(* Logix 5000 project; controller TFF vendor 1 type 14 code 107 rev 34.11; software revision 34.03; part 7 of 36 *)

        [24]   // Product Recovery 1&5 - Empty Recycle Bag (TF3S)
        [16]   // Recycle Bag Fill
        [6]   // Buffer Source Open
        [25]   // Product Recovery 2 - Empty Membranes (TF3S
        [30]   // Filter User
        [34]   // Column User
        [36]   // Fraction 3
        [37]   // Fraction 2
        [61]   // Reserved : Open All valves
        [38]   // Fraction 1
        [18]   // Recovery Filter Flush
        [39]   // System Drain
        [19]   // Batch UF or Membrane Recycle
        [14]   // Membrane Soak
        [2]   // Critical Alarm Flowpath
        [33]   // Column Bypass
        [9]   // Air Source Open
        [4]   // All Source Valves Closed
        [62]   // Reserved : Close All valves
        [3]   // All Source Valves Open
        [8]   // Water Source Open
        [22]   // Product Recovery 2 - Empty Retentate Line (TF2S)
        [26]   // Product Recovery 3&6 - Empty Bypass (TF3S)
        [27]   // Product Recovery 4 - Empty Retentate Line (TF3S)
   FlowPath_Storage : FlowPath[6,64] := ([0,0].Truth1 := -1, [0,0].Mask1 := -1, [0,0].Desc := 'Reserved', [0,1].Status := 1, [0,1].Truth1 := 2097151, [0,1].Mask1 := -1, [0,1].Desc := 'Default', [0,2].Status := 1, [0,2].Truth1 := 539146240, [0,2].Mask1 := -1, [0,2].Desc := 'Critical', [0,3].Status := 1, [0,3].Mask1 := 2047, [0,3].Desc := 'Close All Inlets', [0,4].Truth1 := 17, [0,4].Mask1 := 63, [0,4].Desc := 'Inlet 1A', [0,5].Truth1 := 18, [0,5].Mask1 := 63, [0,5].Desc := 'Inlet 1B', [0,6].Truth1 := 20, [0,6].Mask1 := 63, [0,6].Desc := 'Inlet 1C', [0,7].Truth1 := 24, [0,7].Mask1 := 63, [0,7].Desc := 'Inlet 1D', [0,8].Truth1 := 32, [0,8].Mask1 := 63, [0,8].Desc := 'Inlet 1E', [0,9].Truth1 := 64, [0,9].Mask1 := 1984, [0,9].Desc := 'Inlet 2A', [0,10].Truth1 := 128, [0,10].Mask1 := 1984, [0,10].Desc := 'Inlet 2B', [0,11].Truth1 := 256, [0,11].Mask1 := 1984, [0,11].Desc := 'Inlet 2C', [0,12].Truth1 := 512, [0,12].Mask1 := 1984, [0,12].Desc := 'Inlet 2D', [0,13].Truth1 := 1024, [0,13].Mask1 := 1984, [0,13].Desc := 'Inlet 2E', [0,14].Truth1 := 2047, [0,14].Mask1 := 2047, [0,14].Desc := 'Open All Inlets', [0,15].Truth1 := 2047, [0,15].Mask1 := 2047, [0,15].Desc := 'Flexware Installation', [0,16].Truth1 := 2048, [0,16].Mask1 := -2147477504, [0,16].Desc := 'P001 Process', [0,17].Truth1 := -2147481600, [0,17].Mask1 := -2147477504, [0,17].Desc := 'P001 Drain', [0,18].Truth1 := 4096, [0,18].Mask1 := -2147477504, [0,18].Desc := 'P002 Process', [0,19].Truth1 := -2147479552,
        [0,19].Mask1 := -2147477504, [0,19].Desc := 'P002 Drain', [0,20].Status := 1, [0,20].Truth1 := 6144, [0,20].Mask1 := -2147477504, [0,20].Desc := 'Dual Pumps Process', [0,21].Truth1 := -2147477504, [0,21].Mask1 := -2147477504, [0,21].Desc := 'Dual Pumps Drain', [0,22].Status := 1, [0,22].Truth1 := 40960, [0,22].Mask1 := -1073684480, [0,22].Desc := 'BBT Online', [0,23].Truth1 := 16384, [0,23].Mask1 := -1073684480, [0,23].Desc := 'BBT Bypass', [0,24].Truth1 := 1073741824, [0,24].Mask1 := 1073741824, [0,24].Desc := 'BBT Vent', [0,25].Truth1 := 1073750016, [0,25].Mask1 := -1073684480, [0,25].Desc := 'BBT Clean', [0,26].Truth1 := -1073692672, [0,26].Mask1 := -1073684480, [0,26].Desc := 'BBT Drain', [0,27].Mask1 := -1, [0,27].Desc := 'BBT User', [0,28].Truth1 := 327680, [0,28].Mask1 := 458752, [0,28].Desc := 'Filter Online', [0,29].Status := 1, [0,29].Truth1 := 131072, [0,29].Mask1 := 458752, [0,29].Desc := 'Filter Bypass', [0,30].Mask1 := -1, [0,30].Desc := 'Filter User', [0,31].Truth1 := 59244544, [0,31].Mask1 := 66584576, [0,31].Desc := 'Column Forward', [0,32].Truth1 := 55574528, [0,32].Mask1 := 66584576, [0,32].Desc := 'Column Reverse', [0,33].Status := 1, [0,33].Truth1 := 2097152, [0,33].Mask1 := 66584576, [0,33].Desc := 'Column Bypass', [0,34].Mask1 := -1, [0,34].Desc := 'Column user', [0,35].Status := 1, [0,35].Truth1 := 536870912, [0,35].Mask1 := 1006632960, [0,35].Desc := 'Fraction Waste', [0,36].Truth1 := 268435456, [0,36].Mask1 := 1006632960, [0,36].Desc := 'Fraction 3', [0,37].Truth1 := 134217728, [0,37].Mask1 := 1006632960, [0,37].Desc := 'Fraction 2', [0,38].Truth1 := 67108864, [0,38].Mask1 := 1006632960,
        [0,38].Desc := 'Fraction 1', [0,39].Truth1 := -1, [0,39].Mask1 := -1, [0,39].Desc := 'System Drain', [0,40].Status := 1, [0,40].Desc := 'User 1', [0,41].Status := 1, [0,41].Desc := 'User 2', [0,42].Truth2 := 32768, [0,42].Mask2 := 32960, [0,42].Desc := 'User 3', [0,43].Status := 1, [0,43].Desc := 'User 4', [0,44].Truth1 := 118489088, [0,44].Mask1 := 133169152, [0,44].Desc := 'User 5', [0,45].Status := 1, [0,46].Status := 1, [0,47].Status := 1, [0,48].Status := 1, [0,49].Status := 1, [0,50].Status := 1, [0,51].Status := 1, [0,52].Status := 1, [0,53].Status := 1, [0,54].Status := 1, [0,55].Status := 1, [0,56].Status := 1, [0,57].Status := 1, [0,58].Status := 1, [0,59].Status := 1, [0,60].Status := 1, [0,61].Truth1 := -1, [0,61].Mask1 := -1, [0,62].Mask1 := -1, [0,63].Status := 1, [0,63].Truth1 := 539146240, [0,63].Mask1 := -1, [0,63].Mask2 := -1, [0,63].Mask3 := -1, [0,63].Mask4 := -1, [1,0].FlushTruth := 1, [1,0].DrainTruth := 1, [1,0].FlushMask := 1, [1,0].DrainMask := 1, [1,0].Truth1 := 28735, [1,0].Mask1 := 28735, [1,0].Desc := 'Reserved', [1,1].FlushMask := 1, [1,1].DrainMask := 1, [1,1].Truth1 := 524299, [1,1].Mask1 := 2097151, [1,1].Desc := 'Default', [1,2].Status := 1, [1,2].FlushMask := 1, [1,2].DrainMask := 1, [1,2].Truth1 := 524299, [1,2].Mask1 := 32767, [1,2].Desc := 'Critical', [1,3].Truth1 := 1052608,
        [1,3].Mask1 := 4032, [1,3].Desc := 'All Source Valves Open', [1,4].Status := 1, [1,4].Mask1 := 4032, [1,4].Desc := 'All Source Valves Closed', [1,5].Truth1 := 256, [1,5].Mask1 := 4032, [1,5].Desc := 'Feed Source Open', [1,6].Truth1 := 576, [1,6].Mask1 := 4032, [1,6].Desc := 'Buffer Source Open', [1,7].Truth1 := 1088, [1,7].Mask1 := 4032, [1,7].Desc := 'Caustic Source Open', [1,8].Truth1 := 2112, [1,8].Mask1 := 4032, [1,8].Desc := 'Water Source Open', [1,9].Truth1 := 192, [1,9].Mask1 := 4032, [1,9].Desc := 'Air Source Open', [1,10].FlushTruth := 1, [1,10].DrainTruth := 1, [1,10].FlushMask := 1, [1,10].DrainMask := 1, [1,10].Truth1 := 393227, [1,10].Mask1 := 28735, [1,10].Desc := 'Single Pass Flush (from inlet manifold)', [1,11].DrainTruth := 1, [1,11].FlushMask := 1, [1,11].DrainMask := 1, [1,11].Truth1 := 65547, [1,11].Mask1 := 28735, [1,11].Desc := 'Single Pass Flush (from recycle bag)', [1,12].FlushTruth := 1, [1,12].DrainTruth := 1, [1,12].FlushMask := 1, [1,12].DrainMask := 1, [1,12].Truth1 := 409647, [1,12].Mask1 := 28735, [1,12].Desc := 'System Drain (without recycle bag)', [1,13].DrainTruth := 1, [1,13].FlushMask := 1, [1,13].DrainMask := 1, [1,13].Truth1 := 81983, [1,13].Mask1 := 28735, [1,13].Desc := 'System Drain (from recycle bag)', [1,14].FlushMask := 1, [1,14].DrainMask := 1, [1,14].Truth1 := 65539, [1,14].Mask1 := 28735, [1,14].Desc := 'Membrane Soak', [1,15].FlushMask := 1, [1,15].DrainMask := 1, [1,15].Truth1 := 48, [1,15].Mask1 := 28735, [1,15].Desc := 'Integrity Test', [1,16].FlushMask := 1, [1,16].DrainMask := 1, [1,16].Truth1 := 524312, [1,16].Mask1 := 28735,
        [1,16].Desc := 'Recycle Bag Fill', [1,17].FlushMask := 1, [1,17].DrainMask := 1, [1,17].Truth1 := 81925, [1,17].Mask1 := 28735, [1,17].Desc := 'Recycle Bag Drain', [1,18].FlushMask := 1, [1,18].DrainMask := 1, [1,18].Truth1 := 65541, [1,18].Mask1 := 28735, [1,18].Desc := 'Recovery Filter Flush', [1,19].Status := 1, [1,19].FlushMask := 1, [1,19].DrainMask := 1, [1,19].Truth1 := 589835, [1,19].Mask1 := 28735, [1,19].Desc := 'Batch UF or Membrane Recycle', [1,20].FlushMask := 1, [1,20].DrainMask := 1, [1,20].Truth1 := 589851, [1,20].Mask1 := 28735, [1,20].Desc := 'Fed Batch UF or Diafiltration', [1,21].FlushMask := 1, [1,21].DrainMask := 1, [1,21].Truth1 := 65541, [1,21].Mask1 := 16447, [1,21].Desc := 'Product Recovery 1&3 - Empty Recycle Bag (TF2S)', [1,22].FlushMask := 1, [1,22].DrainMask := 1, [1,22].Truth1 := 524312, [1,22].Mask1 := 16447, [1,22].Desc := 'Product Recovery 2 - Empty Retentate Line (TF2S)', [1,23].FlushMask := 1, [1,23].DrainMask := 1, [1,23].Truth1 := 22, [1,23].Mask1 := 16447, [1,23].Desc := 'Product Recovery 4 - Empty Membranes (TF2S)', [1,24].FlushMask := 1, [1,24].DrainMask := 1, [1,24].Truth1 := 65541, [1,24].Mask1 := 28735, [1,24].Desc := 'Product Recovery 1&5 - Empty Recycle Bag (TF3S)', [1,25].FlushMask := 1, [1,25].DrainMask := 1, [1,25].Truth1 := 22, [1,25].Mask1 := 28735, [1,25].Desc := 'Product Recovery 2 - Empty Membranes (TF3S', [1,26].FlushMask := 1, [1,26].DrainMask := 1, [1,26].Truth1 := 12310, [1,26].Mask1 := 28735, [1,26].Desc := 'Product Recovery 3&6 - Empty Bypass (TF3S)', [1,27].FlushMask := 1, [1,27].DrainMask := 1, [1,27].Truth1 := 524312, [1,27].Mask1 := 28735, [1,27].Desc := 'Product Recovery 4 - Empty Retentate Line (TF3S)', [1,28].FlushMask := 1, [1,28].DrainMask := 1, [1,28].Truth1 := 606271,
        [1,28].Mask1 := 28735, [1,28].Desc := 'All Main Flowpath Valves Open', [1,29].FlushMask := 1, [1,29].DrainMask := 1, [1,29].Mask1 := 28735, [1,29].Desc := 'All Main Flowpath Valves Closed', [1,30].Mask1 := -1, [1,30].Desc := 'Filter User', [1,31].Truth1 := 59244544, [1,31].Mask1 := 66584576, [1,31].Desc := 'Column Forward', [1,32].Truth1 := 55574528, [1,32].Mask1 := 66584576, [1,32].Desc := 'Column Reverse', [1,33].Truth1 := 2097152, [1,33].Mask1 := 66584576, [1,33].Desc := 'Column Bypass', [1,34].Mask1 := -1, [1,34].Desc := 'Column user', [1,35].Truth1 := 2068416, [1,35].Mask1 := 4032, [1,35].Desc := 'Fraction Waste', [1,36].Status := 1, [1,36].Desc := 'Fraction 3', [1,37].Status := 1, [1,37].Desc := 'Fraction 2', [1,38].Status := 1, [1,38].Desc := 'Fraction 1', [1,39].Status := 1, [1,39].Desc := 'System Drain', [1,40].Status := 1, [1,40].Desc := 'User 1', [1,41].Status := 1, [1,41].Desc := 'User 2', [1,42].Status := 1, [1,42].Desc := 'User 3', [1,43].Status := 1, [1,43].Desc := 'User 4', [1,44].Status := 1, [1,44].Desc := 'User 5', [1,45].Status := 1, [1,46].Status := 1, [1,47].Status := 1, [1,48].Status := 1, [1,49].Status := 1, [1,50].Status := 1, [1,51].Status := 1, [1,52].Status := 1, [1,53].Status := 1, [1,54].Status := 1, [1,55].Status := 1, [1,56].Status := 1, [1,57].Status := 1, [1,58].Status := 1, [1,59].Status := 1, [1,60].Status := 1, [1,61].Truth1 := -1, [1,61].Mask1 := -1, [1,62].Mask1 := -1, [1,63].Status := 1,
        [1,63].FlushMask := 1, [1,63].DrainMask := 1, [1,63].Truth1 := 11, [1,63].Mask1 := -1, [1,63].Mask2 := -1, [1,63].Mask3 := -1, [1,63].Mask4 := -1, [2,0].Truth1 := -1, [2,0].Mask1 := -1, [2,0].Desc := 'Reserved', [2,1].Status := 1, [2,1].FlushMask := 1, [2,1].DrainMask := 1, [2,1].Truth1 := 11, [2,1].Mask1 := 2097151, [2,1].Desc := 'Default', [2,2].Status := 1, [2,2].FlushMask := 1, [2,2].DrainMask := 1, [2,2].Truth1 := 11, [2,2].Mask1 := 28735, [2,2].Desc := 'Critical', [2,3].Truth1 := 4032, [2,3].Mask1 := 4032, [2,3].Desc := 'Close All Inlets', [2,4].Status := 1, [2,4].Mask1 := 4032, [2,4].Desc := 'Inlet 1A', [2,5].Truth1 := 256, [2,5].Mask1 := 4032, [2,5].Desc := 'Inlet 1B', [2,6].Truth1 := 576, [2,6].Mask1 := 4032, [2,6].Desc := 'Inlet 1C', [2,7].Truth1 := 1088, [2,7].Mask1 := 4032, [2,7].Desc := 'Inlet 1D', [2,8].Truth1 := 2112, [2,8].Mask1 := 4032, [2,8].Desc := 'Inlet 1E', [2,9].Truth1 := 192, [2,9].Mask1 := 4032, [2,9].Desc := 'Inlet 2A', [2,10].FlushTruth := 1, [2,10].DrainTruth := 1, [2,10].FlushMask := 1, [2,10].DrainMask := 1, [2,10].Truth1 := 11, [2,10].Mask1 := 28735, [2,10].Desc := 'Inlet 2B', [2,11].DrainTruth := 1, [2,11].FlushMask := 1, [2,11].DrainMask := 1, [2,11].Truth1 := 11, [2,11].Mask1 := 28735, [2,11].Desc := 'Inlet 2C', [2,12].FlushTruth := 1, [2,12].DrainTruth := 1, [2,12].FlushMask := 1, [2,12].DrainMask := 1,
        [2,12].Truth1 := 16431, [2,12].Mask1 := 28735, [2,12].Desc := 'Inlet 2D', [2,13].DrainTruth := 1, [2,13].FlushMask := 1, [2,13].DrainMask := 1, [2,13].Truth1 := 16447, [2,13].Mask1 := 28735, [2,13].Desc := 'Inlet 2E', [2,14].FlushMask := 1, [2,14].DrainMask := 1, [2,14].Truth1 := 3, [2,14].Mask1 := 28735, [2,14].Desc := 'Open All Inlets', [2,15].FlushMask := 1, [2,15].DrainMask := 1, [2,15].Truth1 := 48, [2,15].Mask1 := 28735, [2,15].Desc := 'Flexware Installation', [2,16].FlushMask := 1, [2,16].DrainMask := 1, [2,16].Truth1 := 24, [2,16].Mask1 := 28735, [2,16].Desc := 'P001 Process', [2,17].FlushMask := 1, [2,17].DrainMask := 1, [2,17].Truth1 := 16389, [2,17].Mask1 := 28735, [2,17].Desc := 'P001 Drain', [2,18].FlushMask := 1, [2,18].DrainMask := 1, [2,18].Truth1 := 5, [2,18].Mask1 := 28735, [2,18].Desc := 'P002 Process', [2,19].Status := 1, [2,19].FlushMask := 1, [2,19].DrainMask := 1, [2,19].Truth1 := 11, [2,19].Mask1 := 28735, [2,19].Desc := 'P002 Drain', [2,20].FlushMask := 1, [2,20].DrainMask := 1, [2,20].Truth1 := 27, [2,20].Mask1 := 28735, [2,20].Desc := 'Dual Pumps Process', [2,21].FlushMask := 1, [2,21].DrainMask := 1, [2,21].Truth1 := 5, [2,21].Mask1 := 16447, [2,21].Desc := 'Dual Pumps Drain', [2,22].FlushMask := 1, [2,22].DrainMask := 1, [2,22].Truth1 := 24, [2,22].Mask1 := 16447, [2,22].Desc := 'BBT Online', [2,23].FlushMask := 1, [2,23].DrainMask := 1, [2,23].Truth1 := 22, [2,23].Mask1 := 16447, [2,23].Desc := 'BBT Bypass',
        [2,24].FlushMask := 1, [2,24].DrainMask := 1, [2,24].Truth1 := 5, [2,24].Mask1 := 28735, [2,24].Desc := 'BBT Vent', [2,25].FlushMask := 1, [2,25].DrainMask := 1, [2,25].Truth1 := 22, [2,25].Mask1 := 28735, [2,25].Desc := 'BBT Clean', [2,26].FlushMask := 1, [2,26].DrainMask := 1, [2,26].Truth1 := 12310, [2,26].Mask1 := 28735, [2,26].Desc := 'BBT Drain', [2,27].FlushMask := 1, [2,27].DrainMask := 1, [2,27].Truth1 := 24, [2,27].Mask1 := 28735, [2,27].Desc := 'BBT User', [2,28].FlushMask := 1, [2,28].DrainMask := 1, [2,28].Truth1 := 16447, [2,28].Mask1 := 28735, [2,28].Desc := 'Filter Online', [2,29].FlushMask := 1, [2,29].DrainMask := 1, [2,29].Mask1 := 28735, [2,29].Desc := 'Filter Bypass', [2,30].Mask1 := -1, [2,30].Desc := 'Filter User', [2,31].Truth1 := 59244544, [2,31].Mask1 := 66584576, [2,31].Desc := 'Column Forward', [2,32].Truth1 := 55574528, [2,32].Mask1 := 66584576, [2,32].Desc := 'Column Reverse', [2,33].Truth1 := 2097152, [2,33].Mask1 := 66584576, [2,33].Desc := 'Column Bypass', [2,34].Mask1 := -1, [2,34].Desc := 'Column user', [2,35].Status := 1, [2,35].Desc := 'Fraction Waste', [2,36].Status := 1, [2,36].Desc := 'Fraction 3', [2,37].Status := 1, [2,37].Desc := 'Fraction 2', [2,38].Status := 1, [2,38].Desc := 'Fraction 1', [2,39].Status := 1, [2,39].Desc := 'System Drain', [2,40].Status := 1, [2,40].Desc := 'User 1', [2,41].Status := 1, [2,41].Desc := 'User 2', [2,42].Status := 1, [2,42].Desc := 'User 3', [2,43].Status := 1, [2,43].Desc := 'User 4',
        [2,44].Status := 1, [2,44].Desc := 'User 5', [2,45].Status := 1, [2,46].Status := 1, [2,47].Status := 1, [2,48].Status := 1, [2,49].Status := 1, [2,50].Status := 1, [2,51].Status := 1, [2,52].Status := 1, [2,53].Status := 1, [2,54].Status := 1, [2,55].Status := 1, [2,56].Status := 1, [2,57].Status := 1, [2,58].Status := 1, [2,59].Status := 1, [2,60].Status := 1, [2,61].Truth1 := -1, [2,61].Mask1 := -1, [2,62].Mask1 := -1, [2,63].Status := 1, [2,63].FlushMask := 1, [2,63].DrainMask := 1, [2,63].Truth1 := 11, [2,63].Mask1 := -1, [2,63].Mask2 := -1, [2,63].Mask3 := -1, [2,63].Mask4 := -1, [3,0].Status := 1, [3,1].Status := 1, [3,2].Truth1 := 539146240, [3,2].Mask1 := -1, [3,3].Status := 1, [3,3].Mask1 := 2047, [3,4].Truth1 := 17, [3,4].Mask1 := 63, [3,5].Truth1 := 18, [3,5].Mask1 := 63, [3,6].Truth1 := 20, [3,6].Mask1 := 63, [3,7].Truth1 := 24, [3,7].Mask1 := 63, [3,8].Truth1 := 32, [3,8].Mask1 := 63, [3,9].Truth1 := 64, [3,9].Mask1 := 1984, [3,10].Truth1 := 128, [3,10].Mask1 := 1984, [3,11].Truth1 := 256, [3,11].Mask1 := 1984, [3,12].Truth1 := 512, [3,12].Mask1 := 1984, [3,13].Truth1 := 1024, [3,13].Mask1 := 1984, [3,14].Truth1 := 2047, [3,14].Mask1 := 2047, [3,15].Truth1 := 2047, [3,15].Mask1 := 2047, [3,16].Truth1 := 2048,
        [3,16].Mask1 := -2147477504, [3,17].Truth1 := -2147481600, [3,17].Mask1 := -2147477504, [3,18].Truth1 := 4096, [3,18].Mask1 := -2147477504, [3,19].Truth1 := -2147479552, [3,19].Mask1 := -2147477504, [3,20].Truth1 := 6144, [3,20].Mask1 := -2147477504, [3,21].Truth1 := -2147477504, [3,21].Mask1 := -2147477504, [3,22].Truth1 := 40960, [3,22].Mask1 := -1073684480, [3,23].Truth1 := 16384, [3,23].Mask1 := -1073684480, [3,24].Truth1 := 1073741824, [3,24].Mask1 := 1073741824, [3,25].Truth1 := 1073750016, [3,25].Mask1 := -1073684480, [3,26].Truth1 := -1073692672, [3,26].Mask1 := -1073684480, [3,27].Status := 1, [3,28].Truth1 := 327680, [3,28].Mask1 := 458752, [3,29].Truth1 := 131072, [3,29].Mask1 := 458752, [3,30].Status := 1, [3,31].Truth1 := 59244544, [3,31].Mask1 := 66584576, [3,32].Truth1 := 55574528, [3,32].Mask1 := 66584576, [3,33].Truth1 := 2097152, [3,33].Mask1 := 66584576, [3,34].Status := 1, [3,35].Truth1 := 536870912, [3,35].Mask1 := 1006632960, [3,36].Truth1 := 268435456, [3,36].Mask1 := 1006632960, [3,37].Truth1 := 134217728, [3,37].Mask1 := 1006632960, [3,38].Truth1 := 67108864, [3,38].Mask1 := 1006632960, [3,39].Truth1 := -1, [3,39].Mask1 := -1, [3,40].Status := 1, [3,41].Status := 1, [3,42].Status := 1, [3,43].Status := 1, [3,44].Status := 1, [3,45].Status := 1, [3,46].Status := 1, [3,47].Status := 1, [3,48].Status := 1, [3,49].Status := 1, [3,50].Status := 1, [3,51].Status := 1, [3,52].Status := 1, [3,53].Status := 1, [3,54].Status := 1, [3,55].Status := 1,
        [3,56].Status := 1, [3,57].Status := 1, [3,58].Status := 1, [3,59].Status := 1, [3,60].Status := 1, [3,61].Truth1 := -1, [3,61].Mask1 := -1, [3,62].Status := 1, [3,62].Mask1 := -1, [3,63].Status := 1, [4,0].Truth1 := -1, [4,0].Mask1 := -1, [4,0].Desc := 'Reserved', [4,1].Status := 1, [4,1].Truth1 := 539146240, [4,1].Mask1 := -1, [4,1].Desc := 'Default', [4,2].Status := 1, [4,2].Truth1 := 539146240, [4,2].Mask1 := -1, [4,2].Desc := 'Critical', [4,3].Status := 1, [4,3].Mask1 := 2047, [4,3].Desc := 'Close All Inlets', [4,4].Truth1 := 17, [4,4].Mask1 := 63, [4,4].Desc := 'Inlet 1A', [4,5].Truth1 := 18, [4,5].Mask1 := 63, [4,5].Desc := 'Inlet 1B', [4,6].Truth1 := 20, [4,6].Mask1 := 63, [4,6].Desc := 'Inlet 1C', [4,7].Truth1 := 24, [4,7].Mask1 := 63, [4,7].Desc := 'Inlet 1D', [4,8].Truth1 := 32, [4,8].Mask1 := 63, [4,8].Desc := 'Inlet 1E', [4,9].Truth1 := 64, [4,9].Mask1 := 1984, [4,9].Desc := 'Inlet 2A', [4,10].Truth1 := 128, [4,10].Mask1 := 1984, [4,10].Desc := 'Inlet 2B', [4,11].Truth1 := 256, [4,11].Mask1 := 1984, [4,11].Desc := 'Inlet 2C', [4,12].Truth1 := 512, [4,12].Mask1 := 1984, [4,12].Desc := 'Inlet 2D', [4,13].Truth1 := 1024, [4,13].Mask1 := 1984, [4,13].Desc := 'Inlet 2E', [4,14].Truth1 := 2047, [4,14].Mask1 := 2047, [4,14].Desc := 'Open All Inlets', [4,15].Truth1 := 2047, [4,15].Mask1 := 2047, [4,15].Desc := 'Flexware Installation',
        [4,16].Truth1 := 4096, [4,16].Mask1 := -2147477504, [4,16].Desc := 'P001 Process', [4,17].Truth1 := -2147479552, [4,17].Mask1 := -2147477504, [4,17].Desc := 'P001 Drain', [4,18].Truth1 := 2048, [4,18].Mask1 := -2147477504, [4,18].Desc := 'P002 Process', [4,19].Truth1 := -2147481600, [4,19].Mask1 := -2147477504, [4,19].Desc := 'P002 Drain', [4,20].Status := 1, [4,20].Truth1 := 6144, [4,20].Mask1 := -2147477504, [4,20].Desc := 'Dual Pumps Process', [4,21].Truth1 := -2147477504, [4,21].Mask1 := -2147477504, [4,21].Desc := 'Dual Pumps Drain', [4,22].Status := 1, [4,22].Truth1 := 40960, [4,22].Mask1 := -1073684480, [4,22].Desc := 'BBT Online', [4,23].Truth1 := 16384, [4,23].Mask1 := -1073684480, [4,23].Desc := 'BBT Bypass', [4,24].Truth1 := 1073741824, [4,24].Mask1 := 1073741824, [4,24].Desc := 'BBT Vent', [4,25].Truth1 := 1073750016, [4,25].Mask1 := -1073684480, [4,25].Desc := 'BBT Clean', [4,26].Truth1 := -1073692672, [4,26].Mask1 := -1073684480, [4,26].Desc := 'BBT Drain', [4,27].Mask1 := -1, [4,27].Desc := 'BBT User', [4,28].Truth1 := 327680, [4,28].Mask1 := 458752, [4,28].Desc := 'Filter Online', [4,29].Status := 1, [4,29].Truth1 := 131072, [4,29].Mask1 := 458752, [4,29].Desc := 'Filter Bypass', [4,30].Mask1 := -1, [4,30].Desc := 'Filter User', [4,31].Truth1 := 59244544, [4,31].Mask1 := 66584576, [4,31].Desc := 'Column Forward', [4,32].Truth1 := 55574528, [4,32].Mask1 := 66584576, [4,32].Desc := 'Column Reverse', [4,33].Status := 1, [4,33].Truth1 := 2097152, [4,33].Mask1 := 66584576, [4,33].Desc := 'Column Bypass', [4,34].Mask1 := -1, [4,34].Desc := 'Column user', [4,35].Status := 1, [4,35].Truth1 := 536870912,
        [4,35].Mask1 := 1006632960, [4,35].Desc := 'Fraction Waste', [4,36].Truth1 := 268435456, [4,36].Mask1 := 1006632960, [4,36].Desc := 'Fraction 3', [4,37].Truth1 := 134217728, [4,37].Mask1 := 1006632960, [4,37].Desc := 'Fraction 2', [4,38].Truth1 := 67108864, [4,38].Mask1 := 1006632960, [4,38].Desc := 'Fraction 1', [4,39].Truth1 := -1, [4,39].Mask1 := -1, [4,39].Desc := 'System Drain', [4,40].Status := 1, [4,40].Desc := 'User 1', [4,41].Status := 1, [4,41].Desc := 'User 2', [4,42].Truth2 := 32768, [4,42].Mask2 := 32960, [4,42].Desc := 'User 3', [4,43].Status := 1, [4,43].Desc := 'User 4', [4,44].Truth1 := 118489088, [4,44].Mask1 := 133169152, [4,44].Desc := 'User 5', [4,45].Status := 1, [4,46].Status := 1, [4,47].Status := 1, [4,48].Status := 1, [4,49].Status := 1, [4,50].Status := 1, [4,51].Status := 1, [4,52].Status := 1, [4,53].Status := 1, [4,54].Status := 1, [4,55].Status := 1, [4,56].Status := 1, [4,57].Status := 1, [4,58].Status := 1, [4,59].Status := 1, [4,60].Status := 1, [4,61].Truth1 := -1, [4,61].Mask1 := -1, [4,62].Mask1 := -1, [4,63].Status := 1, [4,63].Truth1 := 539146240, [4,63].Mask1 := -1, [4,63].Mask2 := -1, [4,63].Mask3 := -1, [4,63].Mask4 := -1, [5,0].Truth1 := -1, [5,0].Mask1 := -1, [5,0].Desc := 'Reserved', [5,1].Status := 1, [5,1].Truth1 := 539146240, [5,1].Mask1 := -1, [5,1].Desc := 'Default', [5,2].Status := 1, [5,2].Truth1 := 539146240,
        [5,2].Mask1 := -1, [5,2].Desc := 'Critical', [5,3].Status := 1, [5,3].Mask1 := 2047, [5,3].Desc := 'Close All Inlets', [5,4].Truth1 := 17, [5,4].Mask1 := 63, [5,4].Desc := 'Inlet 1A', [5,5].Truth1 := 18, [5,5].Mask1 := 63, [5,5].Desc := 'Inlet 1B', [5,6].Truth1 := 20, [5,6].Mask1 := 63, [5,6].Desc := 'Inlet 1C', [5,7].Truth1 := 24, [5,7].Mask1 := 63, [5,7].Desc := 'Inlet 1D', [5,8].Truth1 := 32, [5,8].Mask1 := 63, [5,8].Desc := 'Inlet 1E', [5,9].Truth1 := 64, [5,9].Mask1 := 1984, [5,9].Desc := 'Inlet 2A', [5,10].Truth1 := 128, [5,10].Mask1 := 1984, [5,10].Desc := 'Inlet 2B', [5,11].Truth1 := 256, [5,11].Mask1 := 1984, [5,11].Desc := 'Inlet 2C', [5,12].Truth1 := 512, [5,12].Mask1 := 1984, [5,12].Desc := 'Inlet 2D', [5,13].Truth1 := 1024, [5,13].Mask1 := 1984, [5,13].Desc := 'Inlet 2E', [5,14].Truth1 := 2047, [5,14].Mask1 := 2047, [5,14].Desc := 'Open All Inlets', [5,15].Truth1 := 2047, [5,15].Mask1 := 2047, [5,15].Desc := 'Flexware Installation', [5,16].Truth1 := 2048, [5,16].Mask1 := -2147477504, [5,16].Desc := 'P001 Process', [5,17].Truth1 := -2147481600, [5,17].Mask1 := -2147477504, [5,17].Desc := 'P001 Drain', [5,18].Truth1 := 4096, [5,18].Mask1 := -2147477504, [5,18].Desc := 'P002 Process', [5,19].Truth1 := -2147479552, [5,19].Mask1 := -2147477504, [5,19].Desc := 'P002 Drain', [5,20].Status := 1, [5,20].Truth1 := 6144, [5,20].Mask1 := -2147477504, [5,20].Desc := 'Dual Pumps Process', [5,21].Truth1 := -2147477504, [5,21].Mask1 := -2147477504, [5,21].Desc := 'Dual Pumps Drain',
        [5,22].Status := 1, [5,22].Truth1 := 40960, [5,22].Mask1 := -1073684480, [5,22].Desc := 'BBT Online', [5,23].Truth1 := 16384, [5,23].Mask1 := -1073684480, [5,23].Desc := 'BBT Bypass', [5,24].Truth1 := 1073741824, [5,24].Mask1 := 1073741824, [5,24].Desc := 'BBT Vent', [5,25].Truth1 := 1073750016, [5,25].Mask1 := -1073684480, [5,25].Desc := 'BBT Clean', [5,26].Truth1 := -1073692672, [5,26].Mask1 := -1073684480, [5,26].Desc := 'BBT Drain', [5,27].Mask1 := -1, [5,27].Desc := 'BBT User', [5,28].Truth1 := 327680, [5,28].Mask1 := 458752, [5,28].Desc := 'Filter Online', [5,29].Status := 1, [5,29].Truth1 := 131072, [5,29].Mask1 := 458752, [5,29].Desc := 'Filter Bypass', [5,30].Mask1 := -1, [5,30].Desc := 'Filter User', [5,31].Truth1 := 59244544, [5,31].Mask1 := 66584576, [5,31].Desc := 'Column Forward', [5,32].Truth1 := 55574528, [5,32].Mask1 := 66584576, [5,32].Desc := 'Column Reverse', [5,33].Status := 1, [5,33].Truth1 := 2097152, [5,33].Mask1 := 66584576, [5,33].Desc := 'Column Bypass', [5,34].Mask1 := -1, [5,34].Desc := 'Column user', [5,35].Status := 1, [5,35].Truth1 := 536870912, [5,35].Mask1 := 1006632960, [5,35].Desc := 'Fraction Waste', [5,36].Truth1 := 268435456, [5,36].Mask1 := 1006632960, [5,36].Desc := 'Fraction 3', [5,37].Truth1 := 134217728, [5,37].Mask1 := 1006632960, [5,37].Desc := 'Fraction 2', [5,38].Truth1 := 67108864, [5,38].Mask1 := 1006632960, [5,38].Desc := 'Fraction 1', [5,39].Truth1 := -1, [5,39].Mask1 := -1, [5,39].Desc := 'System Drain', [5,40].Status := 1, [5,40].Desc := 'User 1', [5,41].Status := 1, [5,41].Desc := 'User 2', [5,42].Truth2 := 32768,
        [5,42].Mask2 := 32960, [5,42].Desc := 'User 3', [5,43].Status := 1, [5,43].Desc := 'User 4', [5,44].Truth1 := 118489088, [5,44].Mask1 := 133169152, [5,44].Desc := 'User 5', [5,45].Status := 1, [5,46].Status := 1, [5,47].Status := 1, [5,48].Status := 1, [5,49].Status := 1, [5,50].Status := 1, [5,51].Status := 1, [5,52].Status := 1, [5,53].Status := 1, [5,54].Status := 1, [5,55].Status := 1, [5,56].Status := 1, [5,57].Status := 1, [5,58].Status := 1, [5,59].Status := 1, [5,60].Status := 1, [5,61].Truth1 := -1, [5,61].Mask1 := -1, [5,62].Mask1 := -1, [5,63].Status := 1, [5,63].Truth1 := 539146240, [5,63].Mask1 := -1, [5,63].Mask2 := -1, [5,63].Mask3 := -1, [5,63].Mask4 := -1);
   FlowPathControl : FlowPathControl := (Valve1 := 18559, MaxFlowPath := 63, Status := 63, StatusHMI := 63, FlowpathEnable[0] := 1, FlowpathEnable[1] := 1, FlowpathEnable[2] := 1, FlowpathEnable[3] := 1, FlowpathEnable[4] := 1, FlowpathEnable[5] := 1, FlowpathEnable[6] := 1, FlowpathEnable[7] := 1, FlowpathEnable[8] := 1, FlowpathEnable[9] := 1, FlowpathEnable[10] := 1, FlowpathEnable[11] := 1, FlowpathEnable[12] := 1, FlowpathEnable[13] := 1, FlowpathEnable[14] := 1, FlowpathEnable[15] := 1, FlowpathEnable[16] := 1, FlowpathEnable[17] := 1, FlowpathEnable[18] := 1, FlowpathEnable[19] := 1, FlowpathEnable[20] := 1, FlowpathEnable[21] := 1, FlowpathEnable[22] := 1, FlowpathEnable[23] := 1, FlowpathEnable[24] := 1, FlowpathEnable[25] := 1, FlowpathEnable[26] := 1, FlowpathEnable[27] := 1, FlowpathEnable[28] := 1, FlowpathEnable[29] := 1, FlowpathEnable[30] := 1, FlowpathEnable[31] := 1, FlowpathEnable[32] := 1, FlowpathEnable[33] := 1, FlowpathEnable[34] := 1, FlowpathEnable[35] := 1, FlowpathEnable[36] := 1, FlowpathEnable[37] := 1, FlowpathEnable[38] := 1, FlowpathEnable[39] := 1, FlowpathEnable[40] := 1, FlowpathEnable[41] := 1, FlowpathEnable[42] := 1, FlowpathEnable[43] := 1, FlowpathEnable[44] := 1, FlowpathEnable[45] := 1, FlowpathEnable[46] := 1, FlowpathEnable[47] := 1, FlowpathEnable[48] := 1, FlowpathEnable[49] := 1, FlowpathEnable[50] := 1, FlowpathEnable[51] := 1, FlowpathEnable[52] := 1, FlowpathEnable[53] := 1, FlowpathEnable[54] := 1, FlowpathEnable[55] := 1,
        FlowpathEnable[56] := 1, FlowpathEnable[57] := 1, FlowpathEnable[58] := 1, FlowpathEnable[59] := 1, FlowpathEnable[60] := 1, FlowpathEnable[61] := 1, FlowpathEnable[62] := 1, FlowpathEnable[63] := 1);   // Flow Path Control
   FlowPathSetup : FlowPathSetup := (Number := 1, Prev := 1);   // Flow Path Setup Data
   FQ_Conc : ALIAS FOR Totalizer[0];   // Concentration Totalizer
   FQ_Diaf : ALIAS FOR Totalizer[1];   // DiafiltrationTotalizer
   GradientLinear : LinearGradient := (Variable := 1, Basis := 1, Y[0] := 50.0);   // (To be keep to avoid error on Recipe Download)
   HoldTime : ALIAS FOR Timers[20];   // Hold Time
   HTCCollectorError : BOOL; {constant}   // Hist. Data Collect. Error
   HTCHeartBeat : BOOL;   // Historical Data Collection heartbeat (Set to 1 by HMI Reset to 0 by PLC)
   LI001 : ALIAS FOR AnalogPoint[44];   // Feed Bag Volume
   LI001Alarm : ALIAS FOR AlarmAnalog[44];   // Feed Bag Volume Alarm
   LogVal : LoggedValue;   // Setpoints to be logged
        .Value[2]   // P001 Linear Velocity setpoint
        .Value[5]   // P002 Linear Velocity setpoint
        .Value[7]   // Mixing Conductivity setpoint
        .Value[6]   // Mixing Percentage setpoint
        .Value[0]   // P001 Manual setpoint
        .Value[3]   // P002 Manual setpoint
        .Value[1]   // P001 Flow setpoint
        .Value[4]   // P002 Flow setpoint
   Membrane_Data : Membrane_Data := (Area := 7.98, Density := 1.0, NWP_TCF := 1.1120849, NWP_TCF_Temp := 20, NWP_TCF_Lookup_25[0] := 2.011, NWP_TCF_Lookup_25[1] := 1.943, NWP_TCF_Lookup_25[2] := 1.879, NWP_TCF_Lookup_25[3] := 1.818, NWP_TCF_Lookup_25[4] := 1.761, NWP_TCF_Lookup_25[5] := 1.706, NWP_TCF_Lookup_25[6] := 1.653, NWP_TCF_Lookup_25[7] := 1.604, NWP_TCF_Lookup_25[8] := 1.556, NWP_TCF_Lookup_25[9] := 1.511, NWP_TCF_Lookup_25[10] := 1.468, NWP_TCF_Lookup_25[11] := 1.426, NWP_TCF_Lookup_25[12] := 1.387, NWP_TCF_Lookup_25[13] := 1.349, NWP_TCF_Lookup_25[14] := 1.313, NWP_TCF_Lookup_25[15] := 1.278, NWP_TCF_Lookup_25[16] := 1.245, NWP_TCF_Lookup_25[17] := 1.213, NWP_TCF_Lookup_25[18] := 1.183, NWP_TCF_Lookup_25[19] := 1.154, NWP_TCF_Lookup_25[20] := 1.126, NWP_TCF_Lookup_25[21] := 1.099, NWP_TCF_Lookup_25[22] := 1.072, NWP_TCF_Lookup_25[23] := 1.047, NWP_TCF_Lookup_25[24] := 1.022, NWP_TCF_Lookup_25[25] := 1.0, NWP_TCF_Lookup_25[26] := 0.978, NWP_TCF_Lookup_25[27] := 0.956, NWP_TCF_Lookup_25[28] := 0.935, NWP_TCF_Lookup_25[29] := 0.915, NWP_TCF_Lookup_25[30] := 0.896, NWP_TCF_Lookup_25[31] := 0.877, NWP_TCF_Lookup_25[32] := 0.859, NWP_TCF_Lookup_25[33] := 0.841, NWP_TCF_Lookup_25[34] := 0.824, NWP_TCF_Lookup_25[35] := 0.808, NWP_TCF_Lookup_25[36] := 0.791, NWP_TCF_Lookup_25[37] := 0.777, NWP_TCF_Lookup_25[38] := 0.761, NWP_TCF_Lookup_25[39] := 0.747, NWP_TCF_Lookup_25[40] := 0.733, NWP_TCF_Lookup_25[41] := 0.719, NWP_TCF_Lookup_25[42] := 0.706, NWP_TCF_Lookup_25[43] := 0.694, NWP_TCF_Lookup_25[44] := 0.681, NWP_TCF_Lookup_25[45] := 0.669, NWP_TCF_Lookup_25[46] := 0.658, NWP_TCF_Lookup_25[47] := 0.646, NWP_TCF_Lookup_25[48] := 0.635, NWP_TCF_Lookup_25[49] := 0.624, NWP_TCF_Lookup_25[50] := 0.614, NWP_TCF_Lookup_25[51] := 0.604, NWP_TCF_Lookup_25[52] := 0.594, AlarmStatus := 1);   // Membrane Data
   Memory_Data : Memory_Data := (Free_Mem_IO := 1024872, Free_Mem_DT := 338240, Free_Memory := 1363112, Total_Mem_IO := 1048576, Total_Mem_DT := 2097152, Total_Memory := 3145728, Biggest_IO_Mem_Size_Ava := 1024528, Biggest_DT_Mem_Size_Ava := 330184, Total_Mem_DT_Real := 2097152.0, Free_Mem_DT_Real := 338240.0, Used_Mem_DT_Real := 1758912.0, Percentage_Used_DT := 83.87146);
   Memory_Message : MESSAGE;   // Data for Message instruction read Memory informations
        MessageParameters(ServiceCode := 16#0003, LocalElement := Memory_Request_Data[0], DestinationTag := Memory_Temp[0], ...)
   Memory_Request_Data : SINT[12] := ([0] := 5, [2] := 1, [4] := 2, [6] := 5, [8] := 6, [10] := 7);   // Source elements for message read Memory informations
   Memory_Temp : INT[29] := ([0] := 5, [1] := 1, [3] := -5926, [4] := 3, [5] := 19024, [6] := 1, [9] := 2, [12] := 4, [14] := 8, [17] := 5, [21] := 6, [23] := -6012, [24] := 3, [25] := 7, [27] := 17010, [28] := 1);   // Destination elements for message read Memory informations
   MiscBOOL : BOOL[64] := ([0] := 1, [1] := 1, [2] := 1, [6] := 1, [9] := 1, [22] := 1, [27] := 1, [28] := 1);   // Misc BOOL Values
   MiscDINT : DINT[32];   // Misc DINT Values
   MiscREAL : REAL[50] := ([35] := 100.0, [36] := 22.0, [37] := 2000.0, [39] := 13.0, [40] := 3000.0, [41] := 30.0, [42] := 48.0);   // Misc Real Values
   MIX001 : ALIAS FOR AnalogPoint[14];   // Mixer Speed
   MIX001_SIG : ALIAS FOR DigitalPoint[104];
   Mixer : Mixer := (Mode := 1, SPManual := 15.0, SPAutoMin := 10.0, SPAutoMax := 50.0, LevelMin := 20.0, LevelMax := 80.0, Alarm_Reset_Cmd_Timer.PRE := 3000);   // Mixer config. structure
   NWP : ALIAS FOR AnalogPoint[45];   // Normalized Water Permeability
   NWPAlarm : ALIAS FOR AlarmAnalog[45];   // NWP Alarm
   OperatingTime : OperatingTime := (DayMax := 30.0, HMICtrl := 1, TimerCtrl.PRE := 10000, CountPre := 2592000, Counter := 9042);
   Operation : Operation[6,251] := ([0,0].Action := 1700001, [0,0].ActionValue := 1.0, [0,1].Step := 1, [0,1].Action := 1700003, [0,1].ActionValue := 1.0, [0,2].Step := 2, [0,2].Action := 1800001, [0,3].Step := 3, [0,3].Action := 1800002, [0,4].Step := 4, [0,4].Action := 2600008, [0,5].Step := 5, [0,5].Action := 2600007, [0,6].Step := 6, [0,6].Action := 2600006, [0,7].Step := 7, [0,7].Action := 2600005, [0,8].Step := 8, [0,8].Action := 2600004, [0,9].Step := 9, [0,9].Action := 2600003, [0,10].Step := 10, [0,10].Action := 2600002, [0,11].Step := 11, [0,11].Action := 2600001, [0,12].Step := 12, [0,12].Action := 2600007, [0,12].ActionValue := 1.0, [0,13].Step := 13, [0,13].Criteria1 := 1100602, [0,13].Criteria1Operator := 1, [0,13].Boolean := 1, [0,13].Criteria2 := 300601, [0,13].Criteria2Operator := 4, [0,13].Action := 2600007, [0,13].Criteria1Value := 60.0, [0,13].Criteria2Value := 1.0, [0,14].Step := 14, [0,14].Criteria1 := 300101, [0,14].Criteria1Operator := 4, [0,14].Action := 700005, [0,14].Criteria1Value := 1.0, [0,14].ActionValue := 10.0, [0,15].Step := 15, [0,15].Action := 800002, [0,15].ActionValue := 1.0, [0,16].Step := 16, [0,16].Criteria1 := 800005, [0,16].Criteria1Operator := 1, [0,16].Action := 700005, [0,16].Criteria1Value := 1.0, [0,16].ActionValue := 4.0, [0,17].Step := 17, [0,17].Action := 700301, [0,17].Label := 10, [0,17].ActionValue := 1.0, [0,18].Step := 18, [0,18].Criteria1 := 1100602, [0,18].Criteria1Operator := 1, [0,18].Boolean := 2,
        [0,18].Criteria2 := 700301, [0,18].Criteria2Operator := 1, [0,18].Action := 2600007, [0,18].Criteria1Value := 2.0, [0,18].ActionValue := 1.0, [0,19].Step := 19, [0,19].Criteria1 := 1100602, [0,19].Criteria1Operator := 1, [0,19].Action := 2600004, [0,19].Criteria1Value := 2.0, [0,19].ActionValue := 1.0, [0,20].Step := 20, [0,20].Criteria1 := 1100602, [0,20].Criteria1Operator := 1, [0,20].Action := 2600002, [0,20].Criteria1Value := 2.0, [0,20].ActionValue := 1.0, [0,21].Step := 21, [0,21].Criteria1 := 1100602, [0,21].Criteria1Operator := 1, [0,21].Boolean := 1, [0,21].Criteria2 := 300601, [0,21].Criteria2Operator := 4, [0,21].Action := 2600004, [0,21].Criteria1Value := 60.0, [0,21].Criteria2Value := 1.0, [0,22].Step := 22, [0,22].Action := 2600002, [0,23].Step := 23, [0,23].Action := 2600007, [0,24].Step := 24, [0,24].Action := 700101, [0,24].ActionValue := 1.0, [0,25].Step := 25, [0,25].Criteria1 := 300601, [0,25].Criteria1Operator := 4, [0,25].Boolean := 2, [0,25].Criteria2 := 300101, [0,25].Criteria2Operator := 4, [0,25].Action := 700005, [0,25].Label := 5, [0,25].Criteria1Value := 1.0, [0,25].Criteria2Value := 1.0, [0,25].ActionValue := 1.0, [0,26].Step := 26, [0,26].Criteria1 := 300101, [0,26].Criteria1Operator := 4, [0,26].Action := 700005, [0,26].ActionValue := 2.0, [0,27].Step := 27, [0,27].Criteria1 := 300601, [0,27].Criteria1Operator := 4, [0,27].Action := 700005, [0,27].ActionValue := 3.0, [0,28].Step := 28, [0,28].Action := 2600003, [0,28].Label := 2, [0,28].ActionValue := 1.0, [0,29].Step := 29, [0,29].Criteria1 := 1100602,
        [0,29].Criteria1Operator := 1, [0,29].Action := 2600003, [0,29].Criteria1Value := 5.0, [0,30].Step := 30, [0,30].Action := 700104, [0,31].Step := 31, [0,31].Action := 800001, [0,31].ActionValue := 1.0, [0,32].Step := 32, [0,32].Criteria1 := 800003, [0,32].Criteria1Operator := 1, [0,32].Boolean := 2, [0,32].Criteria2 := 1100602, [0,32].Criteria2Operator := 1, [0,32].Criteria1Value := 1.0, [0,32].Criteria2Value := 2.0, [0,33].Step := 33, [0,33].Action := 800001, [0,33].ActionValue := 1.0, [0,34].Step := 34, [0,34].Criteria1 := 800003, [0,34].Criteria1Operator := 1, [0,34].Criteria1Value := 1.0, [0,35].Step := 35, [0,35].Criteria1 := 1100602, [0,35].Criteria1Operator := 1, [0,35].Action := 2600004, [0,35].Criteria1Value := 5.0, [0,35].ActionValue := 1.0, [0,36].Step := 36, [0,36].Criteria1 := 1100602, [0,36].Criteria1Operator := 1, [0,36].Action := 2600004, [0,36].Criteria1Value := 5.0, [0,37].Step := 37, [0,37].Criteria1 := 1800001, [0,37].Criteria1Operator := 1, [0,37].Action := 700005, [0,37].ActionValue := 5.0, [0,38].Step := 38, [0,38].Action := 800001, [0,38].ActionValue := 1.0, [0,39].Step := 39, [0,39].Criteria1 := 1100602, [0,39].Criteria1Operator := 1, [0,39].Boolean := 2, [0,39].Criteria2 := 800003, [0,39].Criteria2Operator := 1, [0,39].Action := 700102, [0,39].Criteria1Value := 2.0, [0,39].Criteria2Value := 1.0, [0,39].ActionValue := 1.0, [0,40].Step := 40, [0,40].Action := 700005, [0,40].ActionValue := 4.0, [0,41].Step := 41, [0,41].Action := 800001, [0,41].Label := 3, [0,41].ActionValue := 1.0, [0,42].Step := 42,
        [0,42].Criteria1 := 800003, [0,42].Criteria1Operator := 1, [0,42].Boolean := 2, [0,42].Criteria2 := 1100602, [0,42].Criteria2Operator := 1, [0,42].Action := 2600003, [0,42].Criteria1Value := 1.0, [0,42].Criteria2Value := 2.0, [0,42].ActionValue := 1.0, [0,43].Step := 43, [0,43].Action := 2600001, [0,43].ActionValue := 1.0, [0,44].Step := 44, [0,44].Criteria1 := 1100602, [0,44].Criteria1Operator := 1, [0,44].Action := 800001, [0,44].Criteria1Value := 2.0, [0,44].ActionValue := 1.0, [0,45].Step := 45, [0,45].Criteria1 := 800003, [0,45].Criteria1Operator := 1, [0,45].Boolean := 2, [0,45].Criteria2 := 1100602, [0,45].Criteria2Operator := 1, [0,45].Action := 2600003, [0,45].Criteria1Value := 1.0, [0,45].Criteria2Value := 2.0, [0,46].Step := 46, [0,46].Action := 2600001, [0,47].Step := 47, [0,47].Action := 700005, [0,47].ActionValue := 4.0, [0,48].Step := 48, [0,48].Action := 2600006, [0,48].Label := 1, [0,48].ActionValue := 1.0, [0,49].Step := 49, [0,49].Criteria1 := 1100602, [0,49].Criteria1Operator := 1, [0,49].Action := 2600001, [0,49].Criteria1Value := 2.0, [0,49].ActionValue := 1.0, [0,50].Step := 50, [0,50].Criteria1 := 300601, [0,50].Criteria1Operator := 4, [0,50].Boolean := 2, [0,50].Criteria2 := 300701, [0,50].Criteria2Operator := 4, [0,50].Action := 2600001, [0,51].Step := 51, [0,51].Action := 2600006, [0,52].Step := 52, [0,52].Action := 2600003, [0,52].ActionValue := 1.0, [0,53].Step := 53, [0,53].Criteria1 := 1100602, [0,53].Criteria1Operator := 1, [0,53].Boolean := 2, [0,53].Criteria2 := 300201, [0,53].Criteria2Operator := 4,
        [0,53].Action := 2600003, [0,53].Criteria1Value := 2.0, [0,54].Step := 54, [0,54].Action := 800001, [0,54].ActionValue := 1.0, [0,55].Step := 55, [0,55].Criteria1 := 1100602, [0,55].Criteria1Operator := 1, [0,55].Boolean := 2, [0,55].Criteria2 := 800003, [0,55].Criteria2Operator := 1, [0,55].Criteria1Value := 2.0, [0,55].Criteria2Value := 1.0, [0,56].Step := 56, [0,56].Action := 700401, [0,56].ActionValue := 1.0, [0,57].Step := 57, [0,57].Criteria1 := 700401, [0,57].Criteria1Operator := 1, [0,58].Step := 58, [0,58].Action := 700102, [0,58].Label := 4, [0,58].ActionValue := 1.0, [0,59].Step := 59, [0,59].Action := 700302, [0,59].ActionValue := 1.0, [0,60].Step := 60, [0,60].Criteria1 := 1100602, [0,60].Criteria1Operator := 1, [0,60].Action := 1700011, [0,60].Criteria1Value := 2.0, [0,60].ActionValue := 1.0, [0,61].Criteria1 := -999, [0,61].Criteria1Operator := -999, [0,61].Boolean := -999, [0,61].Criteria2 := -999, [0,61].Criteria2Operator := -999, [0,61].Action := -999, [0,61].Label := -999, [0,61].Criteria1Value := -1000000.0, [0,61].Criteria2Value := -1000000.0, [0,61].ActionValue := -1000000.0, [0,62].Criteria1 := -999, [0,62].Criteria1Operator := -999, [0,62].Boolean := -999, [0,62].Criteria2 := -999, [0,62].Criteria2Operator := -999, [0,62].Action := -999, [0,62].Label := -999, [0,62].Criteria1Value := -1000000.0, [0,62].Criteria2Value := -1000000.0, [0,62].ActionValue := -1000000.0, [0,63].Criteria1 := -999, [0,63].Criteria1Operator := -999, [0,63].Boolean := -999, [0,63].Criteria2 := -999, [0,63].Criteria2Operator := -999, [0,63].Action := -999, [0,63].Label := -999, [0,63].Criteria1Value := -1000000.0,
        [0,63].Criteria2Value := -1000000.0, [0,63].ActionValue := -1000000.0, [0,64].Criteria1 := -999, [0,64].Criteria1Operator := -999, [0,64].Boolean := -999, [0,64].Criteria2 := -999, [0,64].Criteria2Operator := -999, [0,64].Action := -999, [0,64].Label := -999, [0,64].Criteria1Value := -1000000.0, [0,64].Criteria2Value := -1000000.0, [0,64].ActionValue := -1000000.0, [0,65].Criteria1 := -999, [0,65].Criteria1Operator := -999, [0,65].Boolean := -999, [0,65].Criteria2 := -999, [0,65].Criteria2Operator := -999, [0,65].Action := -999, [0,65].Label := -999, [0,65].Criteria1Value := -1000000.0, [0,65].Criteria2Value := -1000000.0, [0,65].ActionValue := -1000000.0, [0,66].Criteria1 := -999, [0,66].Criteria1Operator := -999, [0,66].Boolean := -999, [0,66].Criteria2 := -999, [0,66].Criteria2Operator := -999, [0,66].Action := -999, [0,66].Label := -999, [0,66].Criteria1Value := -1000000.0, [0,66].Criteria2Value := -1000000.0, [0,66].ActionValue := -1000000.0, [0,67].Criteria1 := -999, [0,67].Criteria1Operator := -999, [0,67].Boolean := -999, [0,67].Criteria2 := -999, [0,67].Criteria2Operator := -999, [0,67].Action := -999, [0,67].Label := -999, [0,67].Criteria1Value := -1000000.0, [0,67].Criteria2Value := -1000000.0, [0,67].ActionValue := -1000000.0, [0,68].Criteria1 := -999, [0,68].Criteria1Operator := -999, [0,68].Boolean := -999, [0,68].Criteria2 := -999, [0,68].Criteria2Operator := -999, [0,68].Action := -999, [0,68].Label := -999, [0,68].Criteria1Value := -1000000.0, [0,68].Criteria2Value := -1000000.0, [0,68].ActionValue := -1000000.0, [0,69].Criteria1 := -999, [0,69].Criteria1Operator := -999, [0,69].Boolean := -999, [0,69].Criteria2 := -999, [0,69].Criteria2Operator := -999, [0,69].Action := -999, [0,69].Label := -999, [0,69].Criteria1Value := -1000000.0,
        [0,69].Criteria2Value := -1000000.0, [0,69].ActionValue := -1000000.0, [0,70].Criteria1 := -999, [0,70].Criteria1Operator := -999, [0,70].Boolean := -999, [0,70].Criteria2 := -999, [0,70].Criteria2Operator := -999, [0,70].Action := -999, [0,70].Label := -999, [0,70].Criteria1Value := -1000000.0, [0,70].Criteria2Value := -1000000.0, [0,70].ActionValue := -1000000.0, [0,71].Criteria1 := -999, [0,71].Criteria1Operator := -999, [0,71].Boolean := -999, [0,71].Criteria2 := -999, [0,71].Criteria2Operator := -999, [0,71].Action := -999, [0,71].Label := -999, [0,71].Criteria1Value := -1000000.0, [0,71].Criteria2Value := -1000000.0, [0,71].ActionValue := -1000000.0, [0,72].Criteria1 := -999, [0,72].Criteria1Operator := -999, [0,72].Boolean := -999, [0,72].Criteria2 := -999, [0,72].Criteria2Operator := -999, [0,72].Action := -999, [0,72].Label := -999, [0,72].Criteria1Value := -1000000.0, [0,72].Criteria2Value := -1000000.0, [0,72].ActionValue := -1000000.0, [0,73].Criteria1 := -999, [0,73].Criteria1Operator := -999, [0,73].Boolean := -999, [0,73].Criteria2 := -999, [0,73].Criteria2Operator := -999, [0,73].Action := -999, [0,73].Label := -999, [0,73].Criteria1Value := -1000000.0, [0,73].Criteria2Value := -1000000.0, [0,73].ActionValue := -1000000.0, [0,74].Criteria1 := -999, [0,74].Criteria1Operator := -999, [0,74].Boolean := -999, [0,74].Criteria2 := -999, [0,74].Criteria2Operator := -999, [0,74].Action := -999, [0,74].Label := -999, [0,74].Criteria1Value := -1000000.0, [0,74].Criteria2Value := -1000000.0, [0,74].ActionValue := -1000000.0, [0,75].Criteria1 := -999, [0,75].Criteria1Operator := -999, [0,75].Boolean := -999, [0,75].Criteria2 := -999, [0,75].Criteria2Operator := -999, [0,75].Action := -999, [0,75].Label := -999, [0,75].Criteria1Value := -1000000.0,
        [0,75].Criteria2Value := -1000000.0, [0,75].ActionValue := -1000000.0, [0,76].Criteria1 := -999, [0,76].Criteria1Operator := -999, [0,76].Boolean := -999, [0,76].Criteria2 := -999, [0,76].Criteria2Operator := -999, [0,76].Action := -999, [0,76].Label := -999, [0,76].Criteria1Value := -1000000.0, [0,76].Criteria2Value := -1000000.0, [0,76].ActionValue := -1000000.0, [0,77].Criteria1 := -999, [0,77].Criteria1Operator := -999, [0,77].Boolean := -999, [0,77].Criteria2 := -999, [0,77].Criteria2Operator := -999, [0,77].Action := -999, [0,77].Label := -999, [0,77].Criteria1Value := -1000000.0, [0,77].Criteria2Value := -1000000.0, [0,77].ActionValue := -1000000.0, [0,78].Criteria1 := -999, [0,78].Criteria1Operator := -999, [0,78].Boolean := -999, [0,78].Criteria2 := -999, [0,78].Criteria2Operator := -999, [0,78].Action := -999, [0,78].Label := -999, [0,78].Criteria1Value := -1000000.0, [0,78].Criteria2Value := -1000000.0, [0,78].ActionValue := -1000000.0, [0,79].Criteria1 := -999, [0,79].Criteria1Operator := -999, [0,79].Boolean := -999, [0,79].Criteria2 := -999, [0,79].Criteria2Operator := -999, [0,79].Action := -999, [0,79].Label := -999, [0,79].Criteria1Value := -1000000.0, [0,79].Criteria2Value := -1000000.0, [0,79].ActionValue := -1000000.0, [0,80].Criteria1 := -999, [0,80].Criteria1Operator := -999, [0,80].Boolean := -999, [0,80].Criteria2 := -999, [0,80].Criteria2Operator := -999, [0,80].Action := -999, [0,80].Label := -999, [0,80].Criteria1Value := -1000000.0, [0,80].Criteria2Value := -1000000.0, [0,80].ActionValue := -1000000.0, [0,81].Criteria1 := -999, [0,81].Criteria1Operator := -999, [0,81].Boolean := -999, [0,81].Criteria2 := -999, [0,81].Criteria2Operator := -999, [0,81].Action := -999, [0,81].Label := -999, [0,81].Criteria1Value := -1000000.0,
        [0,81].Criteria2Value := -1000000.0, [0,81].ActionValue := -1000000.0, [0,82].Criteria1 := -999, [0,82].Criteria1Operator := -999, [0,82].Boolean := -999, [0,82].Criteria2 := -999, [0,82].Criteria2Operator := -999, [0,82].Action := -999, [0,82].Label := -999, [0,82].Criteria1Value := -1000000.0, [0,82].Criteria2Value := -1000000.0, [0,82].ActionValue := -1000000.0, [0,83].Criteria1 := -999, [0,83].Criteria1Operator := -999, [0,83].Boolean := -999, [0,83].Criteria2 := -999, [0,83].Criteria2Operator := -999, [0,83].Action := -999, [0,83].Label := -999, [0,83].Criteria1Value := -1000000.0, [0,83].Criteria2Value := -1000000.0, [0,83].ActionValue := -1000000.0, [0,84].Criteria1 := -999, [0,84].Criteria1Operator := -999, [0,84].Boolean := -999, [0,84].Criteria2 := -999, [0,84].Criteria2Operator := -999, [0,84].Action := -999, [0,84].Label := -999, [0,84].Criteria1Value := -1000000.0, [0,84].Criteria2Value := -1000000.0, [0,84].ActionValue := -1000000.0, [0,85].Criteria1 := -999, [0,85].Criteria1Operator := -999, [0,85].Boolean := -999, [0,85].Criteria2 := -999, [0,85].Criteria2Operator := -999, [0,85].Action := -999, [0,85].Label := -999, [0,85].Criteria1Value := -1000000.0, [0,85].Criteria2Value := -1000000.0, [0,85].ActionValue := -1000000.0, [0,86].Criteria1 := -999, [0,86].Criteria1Operator := -999, [0,86].Boolean := -999, [0,86].Criteria2 := -999, [0,86].Criteria2Operator := -999, [0,86].Action := -999, [0,86].Label := -999, [0,86].Criteria1Value := -1000000.0, [0,86].Criteria2Value := -1000000.0, [0,86].ActionValue := -1000000.0, [0,87].Criteria1 := -999, [0,87].Criteria1Operator := -999, [0,87].Boolean := -999, [0,87].Criteria2 := -999, [0,87].Criteria2Operator := -999, [0,87].Action := -999, [0,87].Label := -999, [0,87].Criteria1Value := -1000000.0,
        [0,87].Criteria2Value := -1000000.0, [0,87].ActionValue := -1000000.0, [0,88].Criteria1 := -999, [0,88].Criteria1Operator := -999, [0,88].Boolean := -999, [0,88].Criteria2 := -999, [0,88].Criteria2Operator := -999, [0,88].Action := -999, [0,88].Label := -999, [0,88].Criteria1Value := -1000000.0, [0,88].Criteria2Value := -1000000.0, [0,88].ActionValue := -1000000.0, [0,89].Criteria1 := -999, [0,89].Criteria1Operator := -999, [0,89].Boolean := -999, [0,89].Criteria2 := -999, [0,89].Criteria2Operator := -999, [0,89].Action := -999, [0,89].Label := -999, [0,89].Criteria1Value := -1000000.0, [0,89].Criteria2Value := -1000000.0, [0,89].ActionValue := -1000000.0, [0,90].Criteria1 := -999, [0,90].Criteria1Operator := -999, [0,90].Boolean := -999, [0,90].Criteria2 := -999, [0,90].Criteria2Operator := -999, [0,90].Action := -999, [0,90].Label := -999, [0,90].Criteria1Value := -1000000.0, [0,90].Criteria2Value := -1000000.0, [0,90].ActionValue := -1000000.0, [0,91].Criteria1 := -999, [0,91].Criteria1Operator := -999, [0,91].Boolean := -999, [0,91].Criteria2 := -999, [0,91].Criteria2Operator := -999, [0,91].Action := -999, [0,91].Label := -999, [0,91].Criteria1Value := -1000000.0, [0,91].Criteria2Value := -1000000.0, [0,91].ActionValue := -1000000.0, [0,92].Criteria1 := -999, [0,92].Criteria1Operator := -999, [0,92].Boolean := -999, [0,92].Criteria2 := -999, [0,92].Criteria2Operator := -999, [0,92].Action := -999, [0,92].Label := -999, [0,92].Criteria1Value := -1000000.0, [0,92].Criteria2Value := -1000000.0, [0,92].ActionValue := -1000000.0, [0,93].Criteria1 := -999, [0,93].Criteria1Operator := -999, [0,93].Boolean := -999, [0,93].Criteria2 := -999, [0,93].Criteria2Operator := -999, [0,93].Action := -999, [0,93].Label := -999, [0,93].Criteria1Value := -1000000.0,
        [0,93].Criteria2Value := -1000000.0, [0,93].ActionValue := -1000000.0, [0,94].Criteria1 := -999, [0,94].Criteria1Operator := -999, [0,94].Boolean := -999, [0,94].Criteria2 := -999, [0,94].Criteria2Operator := -999, [0,94].Action := -999, [0,94].Label := -999, [0,94].Criteria1Value := -1000000.0, [0,94].Criteria2Value := -1000000.0, [0,94].ActionValue := -1000000.0, [0,95].Criteria1 := -999, [0,95].Criteria1Operator := -999, [0,95].Boolean := -999, [0,95].Criteria2 := -999, [0,95].Criteria2Operator := -999, [0,95].Action := -999, [0,95].Label := -999, [0,95].Criteria1Value := -1000000.0, [0,95].Criteria2Value := -1000000.0, [0,95].ActionValue := -1000000.0, [0,96].Criteria1 := -999, [0,96].Criteria1Operator := -999, [0,96].Boolean := -999, [0,96].Criteria2 := -999, [0,96].Criteria2Operator := -999, [0,96].Action := -999, [0,96].Label := -999, [0,96].Criteria1Value := -1000000.0, [0,96].Criteria2Value := -1000000.0, [0,96].ActionValue := -1000000.0, [0,97].Criteria1 := -999, [0,97].Criteria1Operator := -999, [0,97].Boolean := -999, [0,97].Criteria2 := -999, [0,97].Criteria2Operator := -999, [0,97].Action := -999, [0,97].Label := -999, [0,97].Criteria1Value := -1000000.0, [0,97].Criteria2Value := -1000000.0, [0,97].ActionValue := -1000000.0, [0,98].Criteria1 := -999, [0,98].Criteria1Operator := -999, [0,98].Boolean := -999, [0,98].Criteria2 := -999, [0,98].Criteria2Operator := -999, [0,98].Action := -999, [0,98].Label := -999, [0,98].Criteria1Value := -1000000.0, [0,98].Criteria2Value := -1000000.0, [0,98].ActionValue := -1000000.0, [0,99].Criteria1 := -999, [0,99].Criteria1Operator := -999, [0,99].Boolean := -999, [0,99].Criteria2 := -999, [0,99].Criteria2Operator := -999, [0,99].Action := -999, [0,99].Label := -999, [0,99].Criteria1Value := -1000000.0,
        [0,99].Criteria2Value := -1000000.0, [0,99].ActionValue := -1000000.0, [0,100].Criteria1 := -999, [0,100].Criteria1Operator := -999, [0,100].Boolean := -999, [0,100].Criteria2 := -999, [0,100].Criteria2Operator := -999, [0,100].Action := -999, [0,100].Label := -999, [0,100].Criteria1Value := -1000000.0, [0,100].Criteria2Value := -1000000.0, [0,100].ActionValue := -1000000.0, [0,101].Criteria1 := -999, [0,101].Criteria1Operator := -999, [0,101].Boolean := -999, [0,101].Criteria2 := -999, [0,101].Criteria2Operator := -999, [0,101].Action := -999, [0,101].Label := -999, [0,101].Criteria1Value := -1000000.0, [0,101].Criteria2Value := -1000000.0, [0,101].ActionValue := -1000000.0, [0,102].Criteria1 := -999, [0,102].Criteria1Operator := -999, [0,102].Boolean := -999, [0,102].Criteria2 := -999, [0,102].Criteria2Operator := -999, [0,102].Action := -999, [0,102].Label := -999, [0,102].Criteria1Value := -1000000.0, [0,102].Criteria2Value := -1000000.0, [0,102].ActionValue := -1000000.0, [0,103].Criteria1 := -999, [0,103].Criteria1Operator := -999, [0,103].Boolean := -999, [0,103].Criteria2 := -999, [0,103].Criteria2Operator := -999, [0,103].Action := -999, [0,103].Label := -999, [0,103].Criteria1Value := -1000000.0, [0,103].Criteria2Value := -1000000.0, [0,103].ActionValue := -1000000.0, [0,104].Criteria1 := -999, [0,104].Criteria1Operator := -999, [0,104].Boolean := -999, [0,104].Criteria2 := -999, [0,104].Criteria2Operator := -999, [0,104].Action := -999, [0,104].Label := -999, [0,104].Criteria1Value := -1000000.0, [0,104].Criteria2Value := -1000000.0, [0,104].ActionValue := -1000000.0, [0,105].Criteria1 := -999, [0,105].Criteria1Operator := -999, [0,105].Boolean := -999, [0,105].Criteria2 := -999, [0,105].Criteria2Operator := -999, [0,105].Action := -999, [0,105].Label := -999, [0,105].Criteria1Value := -1000000.0,
        [0,105].Criteria2Value := -1000000.0, [0,105].ActionValue := -1000000.0, [0,106].Criteria1 := -999, [0,106].Criteria1Operator := -999, [0,106].Boolean := -999, [0,106].Criteria2 := -999, [0,106].Criteria2Operator := -999, [0,106].Action := -999, [0,106].Label := -999, [0,106].Criteria1Value := -1000000.0, [0,106].Criteria2Value := -1000000.0, [0,106].ActionValue := -1000000.0, [0,107].Criteria1 := -999, [0,107].Criteria1Operator := -999, [0,107].Boolean := -999, [0,107].Criteria2 := -999, [0,107].Criteria2Operator := -999, [0,107].Action := -999, [0,107].Label := -999, [0,107].Criteria1Value := -1000000.0, [0,107].Criteria2Value := -1000000.0, [0,107].ActionValue := -1000000.0, [0,108].Criteria1 := -999, [0,108].Criteria1Operator := -999, [0,108].Boolean := -999, [0,108].Criteria2 := -999, [0,108].Criteria2Operator := -999, [0,108].Action := -999, [0,108].Label := -999, [0,108].Criteria1Value := -1000000.0, [0,108].Criteria2Value := -1000000.0, [0,108].ActionValue := -1000000.0, [0,109].Criteria1 := -999, [0,109].Criteria1Operator := -999, [0,109].Boolean := -999, [0,109].Criteria2 := -999, [0,109].Criteria2Operator := -999, [0,109].Action := -999, [0,109].Label := -999, [0,109].Criteria1Value := -1000000.0, [0,109].Criteria2Value := -1000000.0, [0,109].ActionValue := -1000000.0, [0,110].Criteria1 := -999, [0,110].Criteria1Operator := -999, [0,110].Boolean := -999, [0,110].Criteria2 := -999, [0,110].Criteria2Operator := -999, [0,110].Action := -999, [0,110].Label := -999, [0,110].Criteria1Value := -1000000.0, [0,110].Criteria2Value := -1000000.0, [0,110].ActionValue := -1000000.0, [0,111].Criteria1 := -999, [0,111].Criteria1Operator := -999, [0,111].Boolean := -999, [0,111].Criteria2 := -999, [0,111].Criteria2Operator := -999, [0,111].Action := -999, [0,111].Label := -999, [0,111].Criteria1Value := -1000000.0,
        [0,111].Criteria2Value := -1000000.0, [0,111].ActionValue := -1000000.0, [0,112].Criteria1 := -999, [0,112].Criteria1Operator := -999, [0,112].Boolean := -999, [0,112].Criteria2 := -999, [0,112].Criteria2Operator := -999, [0,112].Action := -999, [0,112].Label := -999, [0,112].Criteria1Value := -1000000.0, [0,112].Criteria2Value := -1000000.0, [0,112].ActionValue := -1000000.0, [0,113].Criteria1 := -999, [0,113].Criteria1Operator := -999, [0,113].Boolean := -999, [0,113].Criteria2 := -999, [0,113].Criteria2Operator := -999, [0,113].Action := -999, [0,113].Label := -999, [0,113].Criteria1Value := -1000000.0, [0,113].Criteria2Value := -1000000.0, [0,113].ActionValue := -1000000.0, [0,114].Criteria1 := -999, [0,114].Criteria1Operator := -999, [0,114].Boolean := -999, [0,114].Criteria2 := -999, [0,114].Criteria2Operator := -999, [0,114].Action := -999, [0,114].Label := -999, [0,114].Criteria1Value := -1000000.0, [0,114].Criteria2Value := -1000000.0, [0,114].ActionValue := -1000000.0, [0,115].Criteria1 := -999, [0,115].Criteria1Operator := -999, [0,115].Boolean := -999, [0,115].Criteria2 := -999, [0,115].Criteria2Operator := -999, [0,115].Action := -999, [0,115].Label := -999, [0,115].Criteria1Value := -1000000.0, [0,115].Criteria2Value := -1000000.0, [0,115].ActionValue := -1000000.0, [0,116].Criteria1 := -999, [0,116].Criteria1Operator := -999, [0,116].Boolean := -999, [0,116].Criteria2 := -999, [0,116].Criteria2Operator := -999, [0,116].Action := -999, [0,116].Label := -999, [0,116].Criteria1Value := -1000000.0, [0,116].Criteria2Value := -1000000.0, [0,116].ActionValue := -1000000.0, [0,117].Criteria1 := -999, [0,117].Criteria1Operator := -999, [0,117].Boolean := -999, [0,117].Criteria2 := -999, [0,117].Criteria2Operator := -999, [0,117].Action := -999, [0,117].Label := -999, [0,117].Criteria1Value := -1000000.0,
        [0,117].Criteria2Value := -1000000.0, [0,117].ActionValue := -1000000.0, [0,118].Criteria1 := -999, [0,118].Criteria1Operator := -999, [0,118].Boolean := -999, [0,118].Criteria2 := -999, [0,118].Criteria2Operator := -999, [0,118].Action := -999, [0,118].Label := -999, [0,118].Criteria1Value := -1000000.0, [0,118].Criteria2Value := -1000000.0, [0,118].ActionValue := -1000000.0, [0,119].Criteria1 := -999, [0,119].Criteria1Operator := -999, [0,119].Boolean := -999, [0,119].Criteria2 := -999, [0,119].Criteria2Operator := -999, [0,119].Action := -999, [0,119].Label := -999, [0,119].Criteria1Value := -1000000.0, [0,119].Criteria2Value := -1000000.0, [0,119].ActionValue := -1000000.0, [0,120].Criteria1 := -999, [0,120].Criteria1Operator := -999, [0,120].Boolean := -999, [0,120].Criteria2 := -999, [0,120].Criteria2Operator := -999, [0,120].Action := -999, [0,120].Label := -999, [0,120].Criteria1Value := -1000000.0, [0,120].Criteria2Value := -1000000.0, [0,120].ActionValue := -1000000.0, [0,121].Criteria1 := -999, [0,121].Criteria1Operator := -999, [0,121].Boolean := -999, [0,121].Criteria2 := -999, [0,121].Criteria2Operator := -999, [0,121].Action := -999, [0,121].Label := -999, [0,121].Criteria1Value := -1000000.0, [0,121].Criteria2Value := -1000000.0, [0,121].ActionValue := -1000000.0, [0,122].Criteria1 := -999, [0,122].Criteria1Operator := -999, [0,122].Boolean := -999, [0,122].Criteria2 := -999, [0,122].Criteria2Operator := -999, [0,122].Action := -999, [0,122].Label := -999, [0,122].Criteria1Value := -1000000.0, [0,122].Criteria2Value := -1000000.0, [0,122].ActionValue := -1000000.0, [0,123].Criteria1 := -999, [0,123].Criteria1Operator := -999, [0,123].Boolean := -999, [0,123].Criteria2 := -999, [0,123].Criteria2Operator := -999, [0,123].Action := -999, [0,123].Label := -999, [0,123].Criteria1Value := -1000000.0,
        [0,123].Criteria2Value := -1000000.0, [0,123].ActionValue := -1000000.0, [0,124].Criteria1 := -999, [0,124].Criteria1Operator := -999, [0,124].Boolean := -999, [0,124].Criteria2 := -999, [0,124].Criteria2Operator := -999, [0,124].Action := -999, [0,124].Label := -999, [0,124].Criteria1Value := -1000000.0, [0,124].Criteria2Value := -1000000.0, [0,124].ActionValue := -1000000.0, [0,125].Criteria1 := -999, [0,125].Criteria1Operator := -999, [0,125].Boolean := -999, [0,125].Criteria2 := -999, [0,125].Criteria2Operator := -999, [0,125].Action := -999, [0,125].Label := -999, [0,125].Criteria1Value := -1000000.0, [0,125].Criteria2Value := -1000000.0, [0,125].ActionValue := -1000000.0, [0,126].Criteria1 := -999, [0,126].Criteria1Operator := -999, [0,126].Boolean := -999, [0,126].Criteria2 := -999, [0,126].Criteria2Operator := -999, [0,126].Action := -999, [0,126].Label := -999, [0,126].Criteria1Value := -1000000.0, [0,126].Criteria2Value := -1000000.0, [0,126].ActionValue := -1000000.0, [0,127].Criteria1 := -999, [0,127].Criteria1Operator := -999, [0,127].Boolean := -999, [0,127].Criteria2 := -999, [0,127].Criteria2Operator := -999, [0,127].Action := -999, [0,127].Label := -999, [0,127].Criteria1Value := -1000000.0, [0,127].Criteria2Value := -1000000.0, [0,127].ActionValue := -1000000.0, [0,128].Criteria1 := -999, [0,128].Criteria1Operator := -999, [0,128].Boolean := -999, [0,128].Criteria2 := -999, [0,128].Criteria2Operator := -999, [0,128].Action := -999, [0,128].Label := -999, [0,128].Criteria1Value := -1000000.0, [0,128].Criteria2Value := -1000000.0, [0,128].ActionValue := -1000000.0, [0,129].Criteria1 := -999, [0,129].Criteria1Operator := -999, [0,129].Boolean := -999, [0,129].Criteria2 := -999, [0,129].Criteria2Operator := -999, [0,129].Action := -999, [0,129].Label := -999, [0,129].Criteria1Value := -1000000.0,
        [0,129].Criteria2Value := -1000000.0, [0,129].ActionValue := -1000000.0, [0,130].Criteria1 := -999, [0,130].Criteria1Operator := -999, [0,130].Boolean := -999, [0,130].Criteria2 := -999, [0,130].Criteria2Operator := -999, [0,130].Action := -999, [0,130].Label := -999, [0,130].Criteria1Value := -1000000.0, [0,130].Criteria2Value := -1000000.0, [0,130].ActionValue := -1000000.0, [0,131].Criteria1 := -999, [0,131].Criteria1Operator := -999, [0,131].Boolean := -999, [0,131].Criteria2 := -999, [0,131].Criteria2Operator := -999, [0,131].Action := -999, [0,131].Label := -999, [0,131].Criteria1Value := -1000000.0, [0,131].Criteria2Value := -1000000.0, [0,131].ActionValue := -1000000.0, [0,132].Criteria1 := -999, [0,132].Criteria1Operator := -999, [0,132].Boolean := -999, [0,132].Criteria2 := -999, [0,132].Criteria2Operator := -999, [0,132].Action := -999, [0,132].Label := -999, [0,132].Criteria1Value := -1000000.0, [0,132].Criteria2Value := -1000000.0, [0,132].ActionValue := -1000000.0, [0,133].Criteria1 := -999, [0,133].Criteria1Operator := -999, [0,133].Boolean := -999, [0,133].Criteria2 := -999, [0,133].Criteria2Operator := -999, [0,133].Action := -999, [0,133].Label := -999, [0,133].Criteria1Value := -1000000.0, [0,133].Criteria2Value := -1000000.0, [0,133].ActionValue := -1000000.0, [0,134].Criteria1 := -999, [0,134].Criteria1Operator := -999, [0,134].Boolean := -999, [0,134].Criteria2 := -999, [0,134].Criteria2Operator := -999, [0,134].Action := -999, [0,134].Label := -999, [0,134].Criteria1Value := -1000000.0, [0,134].Criteria2Value := -1000000.0, [0,134].ActionValue := -1000000.0, [0,135].Criteria1 := -999, [0,135].Criteria1Operator := -999, [0,135].Boolean := -999, [0,135].Criteria2 := -999, [0,135].Criteria2Operator := -999, [0,135].Action := -999, [0,135].Label := -999, [0,135].Criteria1Value := -1000000.0,
        [0,135].Criteria2Value := -1000000.0, [0,135].ActionValue := -1000000.0, [0,136].Criteria1 := -999, [0,136].Criteria1Operator := -999, [0,136].Boolean := -999, [0,136].Criteria2 := -999, [0,136].Criteria2Operator := -999, [0,136].Action := -999, [0,136].Label := -999, [0,136].Criteria1Value := -1000000.0, [0,136].Criteria2Value := -1000000.0, [0,136].ActionValue := -1000000.0, [0,137].Criteria1 := -999, [0,137].Criteria1Operator := -999, [0,137].Boolean := -999, [0,137].Criteria2 := -999, [0,137].Criteria2Operator := -999, [0,137].Action := -999, [0,137].Label := -999, [0,137].Criteria1Value := -1000000.0, [0,137].Criteria2Value := -1000000.0, [0,137].ActionValue := -1000000.0, [0,138].Criteria1 := -999, [0,138].Criteria1Operator := -999, [0,138].Boolean := -999, [0,138].Criteria2 := -999, [0,138].Criteria2Operator := -999, [0,138].Action := -999, [0,138].Label := -999, [0,138].Criteria1Value := -1000000.0, [0,138].Criteria2Value := -1000000.0, [0,138].ActionValue := -1000000.0, [0,139].Criteria1 := -999, [0,139].Criteria1Operator := -999, [0,139].Boolean := -999, [0,139].Criteria2 := -999, [0,139].Criteria2Operator := -999, [0,139].Action := -999, [0,139].Label := -999, [0,139].Criteria1Value := -1000000.0, [0,139].Criteria2Value := -1000000.0, [0,139].ActionValue := -1000000.0, [0,140].Criteria1 := -999, [0,140].Criteria1Operator := -999, [0,140].Boolean := -999, [0,140].Criteria2 := -999, [0,140].Criteria2Operator := -999, [0,140].Action := -999, [0,140].Label := -999, [0,140].Criteria1Value := -1000000.0, [0,140].Criteria2Value := -1000000.0, [0,140].ActionValue := -1000000.0, [0,141].Criteria1 := -999, [0,141].Criteria1Operator := -999, [0,141].Boolean := -999, [0,141].Criteria2 := -999, [0,141].Criteria2Operator := -999, [0,141].Action := -999, [0,141].Label := -999, [0,141].Criteria1Value := -1000000.0,
        [0,141].Criteria2Value := -1000000.0, [0,141].ActionValue := -1000000.0, [0,142].Criteria1 := -999, [0,142].Criteria1Operator := -999, [0,142].Boolean := -999, [0,142].Criteria2 := -999, [0,142].Criteria2Operator := -999, [0,142].Action := -999, [0,142].Label := -999, [0,142].Criteria1Value := -1000000.0, [0,142].Criteria2Value := -1000000.0, [0,142].ActionValue := -1000000.0, [0,143].Criteria1 := -999, [0,143].Criteria1Operator := -999, [0,143].Boolean := -999, [0,143].Criteria2 := -999, [0,143].Criteria2Operator := -999, [0,143].Action := -999, [0,143].Label := -999, [0,143].Criteria1Value := -1000000.0, [0,143].Criteria2Value := -1000000.0, [0,143].ActionValue := -1000000.0, [0,144].Criteria1 := -999, [0,144].Criteria1Operator := -999, [0,144].Boolean := -999, [0,144].Criteria2 := -999, [0,144].Criteria2Operator := -999, [0,144].Action := -999, [0,144].Label := -999, [0,144].Criteria1Value := -1000000.0, [0,144].Criteria2Value := -1000000.0, [0,144].ActionValue := -1000000.0, [0,145].Criteria1 := -999, [0,145].Criteria1Operator := -999, [0,145].Boolean := -999, [0,145].Criteria2 := -999, [0,145].Criteria2Operator := -999, [0,145].Action := -999, [0,145].Label := -999, [0,145].Criteria1Value := -1000000.0, [0,145].Criteria2Value := -1000000.0, [0,145].ActionValue := -1000000.0, [0,146].Criteria1 := -999, [0,146].Criteria1Operator := -999, [0,146].Boolean := -999, [0,146].Criteria2 := -999, [0,146].Criteria2Operator := -999, [0,146].Action := -999, [0,146].Label := -999, [0,146].Criteria1Value := -1000000.0, [0,146].Criteria2Value := -1000000.0, [0,146].ActionValue := -1000000.0, [0,147].Criteria1 := -999, [0,147].Criteria1Operator := -999, [0,147].Boolean := -999, [0,147].Criteria2 := -999, [0,147].Criteria2Operator := -999, [0,147].Action := -999, [0,147].Label := -999, [0,147].Criteria1Value := -1000000.0,
        [0,147].Criteria2Value := -1000000.0, [0,147].ActionValue := -1000000.0, [0,148].Criteria1 := -999, [0,148].Criteria1Operator := -999, [0,148].Boolean := -999, [0,148].Criteria2 := -999, [0,148].Criteria2Operator := -999, [0,148].Action := -999, [0,148].Label := -999, [0,148].Criteria1Value := -1000000.0, [0,148].Criteria2Value := -1000000.0, [0,148].ActionValue := -1000000.0, [0,149].Criteria1 := -999, [0,149].Criteria1Operator := -999, [0,149].Boolean := -999, [0,149].Criteria2 := -999, [0,149].Criteria2Operator := -999, [0,149].Action := -999, [0,149].Label := -999, [0,149].Criteria1Value := -1000000.0, [0,149].Criteria2Value := -1000000.0, [0,149].ActionValue := -1000000.0, [0,150].Criteria1 := -999, [0,150].Criteria1Operator := -999, [0,150].Boolean := -999, [0,150].Criteria2 := -999, [0,150].Criteria2Operator := -999, [0,150].Action := -999, [0,150].Label := -999, [0,150].Criteria1Value := -1000000.0, [0,150].Criteria2Value := -1000000.0, [0,150].ActionValue := -1000000.0, [0,151].Criteria1 := -999, [0,151].Criteria1Operator := -999, [0,151].Boolean := -999, [0,151].Criteria2 := -999, [0,151].Criteria2Operator := -999, [0,151].Action := -999, [0,151].Label := -999, [0,151].Criteria1Value := -1000000.0, [0,151].Criteria2Value := -1000000.0, [0,151].ActionValue := -1000000.0, [0,152].Criteria1 := -999, [0,152].Criteria1Operator := -999, [0,152].Boolean := -999, [0,152].Criteria2 := -999, [0,152].Criteria2Operator := -999, [0,152].Action := -999, [0,152].Label := -999, [0,152].Criteria1Value := -1000000.0, [0,152].Criteria2Value := -1000000.0, [0,152].ActionValue := -1000000.0, [0,153].Criteria1 := -999, [0,153].Criteria1Operator := -999, [0,153].Boolean := -999, [0,153].Criteria2 := -999, [0,153].Criteria2Operator := -999, [0,153].Action := -999, [0,153].Label := -999, [0,153].Criteria1Value := -1000000.0,
        [0,153].Criteria2Value := -1000000.0, [0,153].ActionValue := -1000000.0, [0,154].Criteria1 := -999, [0,154].Criteria1Operator := -999, [0,154].Boolean := -999, [0,154].Criteria2 := -999, [0,154].Criteria2Operator := -999, [0,154].Action := -999, [0,154].Label := -999, [0,154].Criteria1Value := -1000000.0, [0,154].Criteria2Value := -1000000.0, [0,154].ActionValue := -1000000.0, [0,155].Criteria1 := -999, [0,155].Criteria1Operator := -999, [0,155].Boolean := -999, [0,155].Criteria2 := -999, [0,155].Criteria2Operator := -999, [0,155].Action := -999, [0,155].Label := -999, [0,155].Criteria1Value := -1000000.0, [0,155].Criteria2Value := -1000000.0, [0,155].ActionValue := -1000000.0, [0,156].Criteria1 := -999, [0,156].Criteria1Operator := -999, [0,156].Boolean := -999, [0,156].Criteria2 := -999, [0,156].Criteria2Operator := -999, [0,156].Action := -999, [0,156].Label := -999, [0,156].Criteria1Value := -1000000.0, [0,156].Criteria2Value := -1000000.0, [0,156].ActionValue := -1000000.0, [0,157].Criteria1 := -999, [0,157].Criteria1Operator := -999, [0,157].Boolean := -999, [0,157].Criteria2 := -999, [0,157].Criteria2Operator := -999, [0,157].Action := -999, [0,157].Label := -999, [0,157].Criteria1Value := -1000000.0, [0,157].Criteria2Value := -1000000.0, [0,157].ActionValue := -1000000.0, [0,158].Criteria1 := -999, [0,158].Criteria1Operator := -999, [0,158].Boolean := -999, [0,158].Criteria2 := -999, [0,158].Criteria2Operator := -999, [0,158].Action := -999, [0,158].Label := -999, [0,158].Criteria1Value := -1000000.0, [0,158].Criteria2Value := -1000000.0, [0,158].ActionValue := -1000000.0, [0,159].Criteria1 := -999, [0,159].Criteria1Operator := -999, [0,159].Boolean := -999, [0,159].Criteria2 := -999, [0,159].Criteria2Operator := -999, [0,159].Action := -999, [0,159].Label := -999, [0,159].Criteria1Value := -1000000.0,
        [0,159].Criteria2Value := -1000000.0, [0,159].ActionValue := -1000000.0, [0,160].Criteria1 := -999, [0,160].Criteria1Operator := -999, [0,160].Boolean := -999, [0,160].Criteria2 := -999, [0,160].Criteria2Operator := -999, [0,160].Action := -999, [0,160].Label := -999, [0,160].Criteria1Value := -1000000.0, [0,160].Criteria2Value := -1000000.0, [0,160].ActionValue := -1000000.0, [0,161].Criteria1 := -999, [0,161].Criteria1Operator := -999, [0,161].Boolean := -999, [0,161].Criteria2 := -999, [0,161].Criteria2Operator := -999, [0,161].Action := -999, [0,161].Label := -999, [0,161].Criteria1Value := -1000000.0, [0,161].Criteria2Value := -1000000.0, [0,161].ActionValue := -1000000.0, [0,162].Criteria1 := -999, [0,162].Criteria1Operator := -999, [0,162].Boolean := -999, [0,162].Criteria2 := -999, [0,162].Criteria2Operator := -999, [0,162].Action := -999, [0,162].Label := -999, [0,162].Criteria1Value := -1000000.0, [0,162].Criteria2Value := -1000000.0, [0,162].ActionValue := -1000000.0, [0,163].Criteria1 := -999, [0,163].Criteria1Operator := -999, [0,163].Boolean := -999, [0,163].Criteria2 := -999, [0,163].Criteria2Operator := -999, [0,163].Action := -999, [0,163].Label := -999, [0,163].Criteria1Value := -1000000.0, [0,163].Criteria2Value := -1000000.0, [0,163].ActionValue := -1000000.0, [0,164].Criteria1 := -999, [0,164].Criteria1Operator := -999, [0,164].Boolean := -999, [0,164].Criteria2 := -999, [0,164].Criteria2Operator := -999, [0,164].Action := -999, [0,164].Label := -999, [0,164].Criteria1Value := -1000000.0, [0,164].Criteria2Value := -1000000.0, [0,164].ActionValue := -1000000.0, [0,165].Criteria1 := -999, [0,165].Criteria1Operator := -999, [0,165].Boolean := -999, [0,165].Criteria2 := -999, [0,165].Criteria2Operator := -999, [0,165].Action := -999, [0,165].Label := -999, [0,165].Criteria1Value := -1000000.0,
        [0,165].Criteria2Value := -1000000.0, [0,165].ActionValue := -1000000.0, [0,166].Criteria1 := -999, [0,166].Criteria1Operator := -999, [0,166].Boolean := -999, [0,166].Criteria2 := -999, [0,166].Criteria2Operator := -999, [0,166].Action := -999, [0,166].Label := -999, [0,166].Criteria1Value := -1000000.0, [0,166].Criteria2Value := -1000000.0, [0,166].ActionValue := -1000000.0, [0,167].Criteria1 := -999, [0,167].Criteria1Operator := -999, [0,167].Boolean := -999, [0,167].Criteria2 := -999, [0,167].Criteria2Operator := -999, [0,167].Action := -999, [0,167].Label := -999, [0,167].Criteria1Value := -1000000.0, [0,167].Criteria2Value := -1000000.0, [0,167].ActionValue := -1000000.0, [0,168].Criteria1 := -999, [0,168].Criteria1Operator := -999, [0,168].Boolean := -999, [0,168].Criteria2 := -999, [0,168].Criteria2Operator := -999, [0,168].Action := -999, [0,168].Label := -999, [0,168].Criteria1Value := -1000000.0, [0,168].Criteria2Value := -1000000.0, [0,168].ActionValue := -1000000.0, [0,169].Criteria1 := -999, [0,169].Criteria1Operator := -999, [0,169].Boolean := -999, [0,169].Criteria2 := -999, [0,169].Criteria2Operator := -999, [0,169].Action := -999, [0,169].Label := -999, [0,169].Criteria1Value := -1000000.0, [0,169].Criteria2Value := -1000000.0, [0,169].ActionValue := -1000000.0, [0,170].Criteria1 := -999, [0,170].Criteria1Operator := -999, [0,170].Boolean := -999, [0,170].Criteria2 := -999, [0,170].Criteria2Operator := -999, [0,170].Action := -999, [0,170].Label := -999, [0,170].Criteria1Value := -1000000.0, [0,170].Criteria2Value := -1000000.0, [0,170].ActionValue := -1000000.0, [0,171].Criteria1 := -999, [0,171].Criteria1Operator := -999, [0,171].Boolean := -999, [0,171].Criteria2 := -999, [0,171].Criteria2Operator := -999, [0,171].Action := -999, [0,171].Label := -999, [0,171].Criteria1Value := -1000000.0,
        [0,171].Criteria2Value := -1000000.0, [0,171].ActionValue := -1000000.0, [0,172].Criteria1 := -999, [0,172].Criteria1Operator := -999, [0,172].Boolean := -999, [0,172].Criteria2 := -999, [0,172].Criteria2Operator := -999, [0,172].Action := -999, [0,172].Label := -999, [0,172].Criteria1Value := -1000000.0, [0,172].Criteria2Value := -1000000.0, [0,172].ActionValue := -1000000.0, [0,173].Criteria1 := -999, [0,173].Criteria1Operator := -999, [0,173].Boolean := -999, [0,173].Criteria2 := -999, [0,173].Criteria2Operator := -999, [0,173].Action := -999, [0,173].Label := -999, [0,173].Criteria1Value := -1000000.0, [0,173].Criteria2Value := -1000000.0, [0,173].ActionValue := -1000000.0, [0,174].Criteria1 := -999, [0,174].Criteria1Operator := -999, [0,174].Boolean := -999, [0,174].Criteria2 := -999, [0,174].Criteria2Operator := -999, [0,174].Action := -999, [0,174].Label := -999, [0,174].Criteria1Value := -1000000.0, [0,174].Criteria2Value := -1000000.0, [0,174].ActionValue := -1000000.0, [0,175].Criteria1 := -999, [0,175].Criteria1Operator := -999, [0,175].Boolean := -999, [0,175].Criteria2 := -999, [0,175].Criteria2Operator := -999, [0,175].Action := -999, [0,175].Label := -999, [0,175].Criteria1Value := -1000000.0, [0,175].Criteria2Value := -1000000.0, [0,175].ActionValue := -1000000.0, [0,176].Criteria1 := -999, [0,176].Criteria1Operator := -999, [0,176].Boolean := -999, [0,176].Criteria2 := -999, [0,176].Criteria2Operator := -999, [0,176].Action := -999, [0,176].Label := -999, [0,176].Criteria1Value := -1000000.0, [0,176].Criteria2Value := -1000000.0, [0,176].ActionValue := -1000000.0, [0,177].Criteria1 := -999, [0,177].Criteria1Operator := -999, [0,177].Boolean := -999, [0,177].Criteria2 := -999, [0,177].Criteria2Operator := -999, [0,177].Action := -999, [0,177].Label := -999, [0,177].Criteria1Value := -1000000.0,
        [0,177].Criteria2Value := -1000000.0, [0,177].ActionValue := -1000000.0, [0,178].Criteria1 := -999, [0,178].Criteria1Operator := -999, [0,178].Boolean := -999, [0,178].Criteria2 := -999, [0,178].Criteria2Operator := -999, [0,178].Action := -999, [0,178].Label := -999, [0,178].Criteria1Value := -1000000.0, [0,178].Criteria2Value := -1000000.0, [0,178].ActionValue := -1000000.0, [0,179].Criteria1 := -999, [0,179].Criteria1Operator := -999, [0,179].Boolean := -999, [0,179].Criteria2 := -999, [0,179].Criteria2Operator := -999, [0,179].Action := -999, [0,179].Label := -999, [0,179].Criteria1Value := -1000000.0, [0,179].Criteria2Value := -1000000.0, [0,179].ActionValue := -1000000.0, [0,180].Criteria1 := -999, [0,180].Criteria1Operator := -999, [0,180].Boolean := -999, [0,180].Criteria2 := -999, [0,180].Criteria2Operator := -999, [0,180].Action := -999, [0,180].Label := -999, [0,180].Criteria1Value := -1000000.0, [0,180].Criteria2Value := -1000000.0, [0,180].ActionValue := -1000000.0, [0,181].Criteria1 := -999, [0,181].Criteria1Operator := -999, [0,181].Boolean := -999, [0,181].Criteria2 := -999, [0,181].Criteria2Operator := -999, [0,181].Action := -999, [0,181].Label := -999, [0,181].Criteria1Value := -1000000.0, [0,181].Criteria2Value := -1000000.0, [0,181].ActionValue := -1000000.0, [0,182].Criteria1 := -999, [0,182].Criteria1Operator := -999, [0,182].Boolean := -999, [0,182].Criteria2 := -999, [0,182].Criteria2Operator := -999, [0,182].Action := -999, [0,182].Label := -999, [0,182].Criteria1Value := -1000000.0, [0,182].Criteria2Value := -1000000.0, [0,182].ActionValue := -1000000.0, [0,183].Criteria1 := -999, [0,183].Criteria1Operator := -999, [0,183].Boolean := -999, [0,183].Criteria2 := -999, [0,183].Criteria2Operator := -999, [0,183].Action := -999, [0,183].Label := -999, [0,183].Criteria1Value := -1000000.0,
        [0,183].Criteria2Value := -1000000.0, [0,183].ActionValue := -1000000.0, [0,184].Criteria1 := -999, [0,184].Criteria1Operator := -999, [0,184].Boolean := -999, [0,184].Criteria2 := -999, [0,184].Criteria2Operator := -999, [0,184].Action := -999, [0,184].Label := -999, [0,184].Criteria1Value := -1000000.0, [0,184].Criteria2Value := -1000000.0, [0,184].ActionValue := -1000000.0, [0,185].Criteria1 := -999, [0,185].Criteria1Operator := -999, [0,185].Boolean := -999, [0,185].Criteria2 := -999, [0,185].Criteria2Operator := -999, [0,185].Action := -999, [0,185].Label := -999, [0,185].Criteria1Value := -1000000.0, [0,185].Criteria2Value := -1000000.0, [0,185].ActionValue := -1000000.0, [0,186].Criteria1 := -999, [0,186].Criteria1Operator := -999, [0,186].Boolean := -999, [0,186].Criteria2 := -999, [0,186].Criteria2Operator := -999, [0,186].Action := -999, [0,186].Label := -999, [0,186].Criteria1Value := -1000000.0, [0,186].Criteria2Value := -1000000.0, [0,186].ActionValue := -1000000.0, [0,187].Criteria1 := -999, [0,187].Criteria1Operator := -999, [0,187].Boolean := -999, [0,187].Criteria2 := -999, [0,187].Criteria2Operator := -999, [0,187].Action := -999, [0,187].Label := -999, [0,187].Criteria1Value := -1000000.0, [0,187].Criteria2Value := -1000000.0, [0,187].ActionValue := -1000000.0, [0,188].Criteria1 := -999, [0,188].Criteria1Operator := -999, [0,188].Boolean := -999, [0,188].Criteria2 := -999, [0,188].Criteria2Operator := -999, [0,188].Action := -999, [0,188].Label := -999, [0,188].Criteria1Value := -1000000.0, [0,188].Criteria2Value := -1000000.0, [0,188].ActionValue := -1000000.0, [0,189].Criteria1 := -999, [0,189].Criteria1Operator := -999, [0,189].Boolean := -999, [0,189].Criteria2 := -999, [0,189].Criteria2Operator := -999, [0,189].Action := -999, [0,189].Label := -999, [0,189].Criteria1Value := -1000000.0,
        [0,189].Criteria2Value := -1000000.0, [0,189].ActionValue := -1000000.0, [0,190].Criteria1 := -999, [0,190].Criteria1Operator := -999, [0,190].Boolean := -999, [0,190].Criteria2 := -999, [0,190].Criteria2Operator := -999, [0,190].Action := -999, [0,190].Label := -999, [0,190].Criteria1Value := -1000000.0, [0,190].Criteria2Value := -1000000.0, [0,190].ActionValue := -1000000.0, [0,191].Criteria1 := -999, [0,191].Criteria1Operator := -999, [0,191].Boolean := -999, [0,191].Criteria2 := -999, [0,191].Criteria2Operator := -999, [0,191].Action := -999, [0,191].Label := -999, [0,191].Criteria1Value := -1000000.0, [0,191].Criteria2Value := -1000000.0, [0,191].ActionValue := -1000000.0, [0,192].Criteria1 := -999, [0,192].Criteria1Operator := -999, [0,192].Boolean := -999, [0,192].Criteria2 := -999, [0,192].Criteria2Operator := -999, [0,192].Action := -999, [0,192].Label := -999, [0,192].Criteria1Value := -1000000.0, [0,192].Criteria2Value := -1000000.0, [0,192].ActionValue := -1000000.0, [0,193].Criteria1 := -999, [0,193].Criteria1Operator := -999, [0,193].Boolean := -999, [0,193].Criteria2 := -999, [0,193].Criteria2Operator := -999, [0,193].Action := -999, [0,193].Label := -999, [0,193].Criteria1Value := -1000000.0, [0,193].Criteria2Value := -1000000.0, [0,193].ActionValue := -1000000.0, [0,194].Criteria1 := -999, [0,194].Criteria1Operator := -999, [0,194].Boolean := -999, [0,194].Criteria2 := -999, [0,194].Criteria2Operator := -999, [0,194].Action := -999, [0,194].Label := -999, [0,194].Criteria1Value := -1000000.0, [0,194].Criteria2Value := -1000000.0, [0,194].ActionValue := -1000000.0, [0,195].Criteria1 := -999, [0,195].Criteria1Operator := -999, [0,195].Boolean := -999, [0,195].Criteria2 := -999, [0,195].Criteria2Operator := -999, [0,195].Action := -999, [0,195].Label := -999, [0,195].Criteria1Value := -1000000.0,
        [0,195].Criteria2Value := -1000000.0, [0,195].ActionValue := -1000000.0, [0,196].Criteria1 := -999, [0,196].Criteria1Operator := -999, [0,196].Boolean := -999, [0,196].Criteria2 := -999, [0,196].Criteria2Operator := -999, [0,196].Action := -999, [0,196].Label := -999, [0,196].Criteria1Value := -1000000.0, [0,196].Criteria2Value := -1000000.0, [0,196].ActionValue := -1000000.0, [0,197].Criteria1 := -999, [0,197].Criteria1Operator := -999, [0,197].Boolean := -999, [0,197].Criteria2 := -999, [0,197].Criteria2Operator := -999, [0,197].Action := -999, [0,197].Label := -999, [0,197].Criteria1Value := -1000000.0, [0,197].Criteria2Value := -1000000.0, [0,197].ActionValue := -1000000.0, [0,198].Criteria1 := -999, [0,198].Criteria1Operator := -999, [0,198].Boolean := -999, [0,198].Criteria2 := -999, [0,198].Criteria2Operator := -999, [0,198].Action := -999, [0,198].Label := -999, [0,198].Criteria1Value := -1000000.0, [0,198].Criteria2Value := -1000000.0, [0,198].ActionValue := -1000000.0, [0,199].Criteria1 := -999, [0,199].Criteria1Operator := -999, [0,199].Boolean := -999, [0,199].Criteria2 := -999, [0,199].Criteria2Operator := -999, [0,199].Action := -999, [0,199].Label := -999, [0,199].Criteria1Value := -1000000.0, [0,199].Criteria2Value := -1000000.0, [0,199].ActionValue := -1000000.0, [0,200].Criteria1 := -999, [0,200].Criteria1Operator := -999, [0,200].Boolean := -999, [0,200].Criteria2 := -999, [0,200].Criteria2Operator := -999, [0,200].Action := -999, [0,200].Label := -999, [0,200].Criteria1Value := -1000000.0, [0,200].Criteria2Value := -1000000.0, [0,200].ActionValue := -1000000.0, [0,201].Criteria1 := -999, [0,201].Criteria1Operator := -999, [0,201].Boolean := -999, [0,201].Criteria2 := -999, [0,201].Criteria2Operator := -999, [0,201].Action := -999, [0,201].Label := -999, [0,201].Criteria1Value := -1000000.0,
        [0,201].Criteria2Value := -1000000.0, [0,201].ActionValue := -1000000.0, [0,202].Criteria1 := -999, [0,202].Criteria1Operator := -999, [0,202].Boolean := -999, [0,202].Criteria2 := -999, [0,202].Criteria2Operator := -999, [0,202].Action := -999, [0,202].Label := -999, [0,202].Criteria1Value := -1000000.0, [0,202].Criteria2Value := -1000000.0, [0,202].ActionValue := -1000000.0, [0,203].Criteria1 := -999, [0,203].Criteria1Operator := -999, [0,203].Boolean := -999, [0,203].Criteria2 := -999, [0,203].Criteria2Operator := -999, [0,203].Action := -999, [0,203].Label := -999, [0,203].Criteria1Value := -1000000.0, [0,203].Criteria2Value := -1000000.0, [0,203].ActionValue := -1000000.0, [0,204].Criteria1 := -999, [0,204].Criteria1Operator := -999, [0,204].Boolean := -999, [0,204].Criteria2 := -999, [0,204].Criteria2Operator := -999, [0,204].Action := -999, [0,204].Label := -999, [0,204].Criteria1Value := -1000000.0, [0,204].Criteria2Value := -1000000.0, [0,204].ActionValue := -1000000.0, [0,205].Criteria1 := -999, [0,205].Criteria1Operator := -999, [0,205].Boolean := -999, [0,205].Criteria2 := -999, [0,205].Criteria2Operator := -999, [0,205].Action := -999, [0,205].Label := -999, [0,205].Criteria1Value := -1000000.0, [0,205].Criteria2Value := -1000000.0, [0,205].ActionValue := -1000000.0, [0,206].Criteria1 := -999, [0,206].Criteria1Operator := -999, [0,206].Boolean := -999, [0,206].Criteria2 := -999, [0,206].Criteria2Operator := -999, [0,206].Action := -999, [0,206].Label := -999, [0,206].Criteria1Value := -1000000.0, [0,206].Criteria2Value := -1000000.0, [0,206].ActionValue := -1000000.0, [0,207].Criteria1 := -999, [0,207].Criteria1Operator := -999, [0,207].Boolean := -999, [0,207].Criteria2 := -999, [0,207].Criteria2Operator := -999, [0,207].Action := -999, [0,207].Label := -999, [0,207].Criteria1Value := -1000000.0,
        [0,207].Criteria2Value := -1000000.0, [0,207].ActionValue := -1000000.0, [0,208].Criteria1 := -999, [0,208].Criteria1Operator := -999, [0,208].Boolean := -999, [0,208].Criteria2 := -999, [0,208].Criteria2Operator := -999, [0,208].Action := -999, [0,208].Label := -999, [0,208].Criteria1Value := -1000000.0, [0,208].Criteria2Value := -1000000.0, [0,208].ActionValue := -1000000.0, [0,209].Criteria1 := -999, [0,209].Criteria1Operator := -999, [0,209].Boolean := -999, [0,209].Criteria2 := -999, [0,209].Criteria2Operator := -999, [0,209].Action := -999, [0,209].Label := -999, [0,209].Criteria1Value := -1000000.0, [0,209].Criteria2Value := -1000000.0, [0,209].ActionValue := -1000000.0, [0,210].Criteria1 := -999, [0,210].Criteria1Operator := -999, [0,210].Boolean := -999, [0,210].Criteria2 := -999, [0,210].Criteria2Operator := -999, [0,210].Action := -999, [0,210].Label := -999, [0,210].Criteria1Value := -1000000.0, [0,210].Criteria2Value := -1000000.0, [0,210].ActionValue := -1000000.0, [0,211].Criteria1 := -999, [0,211].Criteria1Operator := -999, [0,211].Boolean := -999, [0,211].Criteria2 := -999, [0,211].Criteria2Operator := -999, [0,211].Action := -999, [0,211].Label := -999, [0,211].Criteria1Value := -1000000.0, [0,211].Criteria2Value := -1000000.0, [0,211].ActionValue := -1000000.0, [0,212].Criteria1 := -999, [0,212].Criteria1Operator := -999, [0,212].Boolean := -999, [0,212].Criteria2 := -999, [0,212].Criteria2Operator := -999, [0,212].Action := -999, [0,212].Label := -999, [0,212].Criteria1Value := -1000000.0, [0,212].Criteria2Value := -1000000.0, [0,212].ActionValue := -1000000.0, [0,213].Criteria1 := -999, [0,213].Criteria1Operator := -999, [0,213].Boolean := -999, [0,213].Criteria2 := -999, [0,213].Criteria2Operator := -999, [0,213].Action := -999, [0,213].Label := -999, [0,213].Criteria1Value := -1000000.0,
        [0,213].Criteria2Value := -1000000.0, [0,213].ActionValue := -1000000.0, [0,214].Criteria1 := -999, [0,214].Criteria1Operator := -999, [0,214].Boolean := -999, [0,214].Criteria2 := -999, [0,214].Criteria2Operator := -999, [0,214].Action := -999, [0,214].Label := -999, [0,214].Criteria1Value := -1000000.0, [0,214].Criteria2Value := -1000000.0, [0,214].ActionValue := -1000000.0, [0,215].Criteria1 := -999, [0,215].Criteria1Operator := -999, [0,215].Boolean := -999, [0,215].Criteria2 := -999, [0,215].Criteria2Operator := -999, [0,215].Action := -999, [0,215].Label := -999, [0,215].Criteria1Value := -1000000.0, [0,215].Criteria2Value := -1000000.0, [0,215].ActionValue := -1000000.0, [0,216].Criteria1 := -999, [0,216].Criteria1Operator := -999, [0,216].Boolean := -999, [0,216].Criteria2 := -999, [0,216].Criteria2Operator := -999, [0,216].Action := -999, [0,216].Label := -999, [0,216].Criteria1Value := -1000000.0, [0,216].Criteria2Value := -1000000.0, [0,216].ActionValue := -1000000.0, [0,217].Criteria1 := -999, [0,217].Criteria1Operator := -999, [0,217].Boolean := -999, [0,217].Criteria2 := -999, [0,217].Criteria2Operator := -999, [0,217].Action := -999, [0,217].Label := -999, [0,217].Criteria1Value := -1000000.0, [0,217].Criteria2Value := -1000000.0, [0,217].ActionValue := -1000000.0, [0,218].Criteria1 := -999, [0,218].Criteria1Operator := -999, [0,218].Boolean := -999, [0,218].Criteria2 := -999, [0,218].Criteria2Operator := -999, [0,218].Action := -999, [0,218].Label := -999, [0,218].Criteria1Value := -1000000.0, [0,218].Criteria2Value := -1000000.0, [0,218].ActionValue := -1000000.0, [0,219].Criteria1 := -999, [0,219].Criteria1Operator := -999, [0,219].Boolean := -999, [0,219].Criteria2 := -999, [0,219].Criteria2Operator := -999, [0,219].Action := -999, [0,219].Label := -999, [0,219].Criteria1Value := -1000000.0,
        [0,219].Criteria2Value := -1000000.0, [0,219].ActionValue := -1000000.0, [0,220].Criteria1 := -999, [0,220].Criteria1Operator := -999, [0,220].Boolean := -999, [0,220].Criteria2 := -999, [0,220].Criteria2Operator := -999, [0,220].Action := -999, [0,220].Label := -999, [0,220].Criteria1Value := -1000000.0, [0,220].Criteria2Value := -1000000.0, [0,220].ActionValue := -1000000.0, [0,221].Criteria1 := -999, [0,221].Criteria1Operator := -999, [0,221].Boolean := -999, [0,221].Criteria2 := -999, [0,221].Criteria2Operator := -999, [0,221].Action := -999, [0,221].Label := -999, [0,221].Criteria1Value := -1000000.0, [0,221].Criteria2Value := -1000000.0, [0,221].ActionValue := -1000000.0, [0,222].Criteria1 := -999, [0,222].Criteria1Operator := -999, [0,222].Boolean := -999, [0,222].Criteria2 := -999, [0,222].Criteria2Operator := -999, [0,222].Action := -999, [0,222].Label := -999, [0,222].Criteria1Value := -1000000.0, [0,222].Criteria2Value := -1000000.0, [0,222].ActionValue := -1000000.0, [0,223].Criteria1 := -999, [0,223].Criteria1Operator := -999, [0,223].Boolean := -999, [0,223].Criteria2 := -999, [0,223].Criteria2Operator := -999, [0,223].Action := -999, [0,223].Label := -999, [0,223].Criteria1Value := -1000000.0, [0,223].Criteria2Value := -1000000.0, [0,223].ActionValue := -1000000.0, [0,224].Criteria1 := -999, [0,224].Criteria1Operator := -999, [0,224].Boolean := -999, [0,224].Criteria2 := -999, [0,224].Criteria2Operator := -999, [0,224].Action := -999, [0,224].Label := -999, [0,224].Criteria1Value := -1000000.0, [0,224].Criteria2Value := -1000000.0, [0,224].ActionValue := -1000000.0, [0,225].Criteria1 := -999, [0,225].Criteria1Operator := -999, [0,225].Boolean := -999, [0,225].Criteria2 := -999, [0,225].Criteria2Operator := -999, [0,225].Action := -999, [0,225].Label := -999, [0,225].Criteria1Value := -1000000.0,
        [0,225].Criteria2Value := -1000000.0, [0,225].ActionValue := -1000000.0, [0,226].Criteria1 := -999, [0,226].Criteria1Operator := -999, [0,226].Boolean := -999, [0,226].Criteria2 := -999, [0,226].Criteria2Operator := -999, [0,226].Action := -999, [0,226].Label := -999, [0,226].Criteria1Value := -1000000.0, [0,226].Criteria2Value := -1000000.0, [0,226].ActionValue := -1000000.0, [0,227].Criteria1 := -999, [0,227].Criteria1Operator := -999, [0,227].Boolean := -999, [0,227].Criteria2 := -999, [0,227].Criteria2Operator := -999, [0,227].Action := -999, [0,227].Label := -999, [0,227].Criteria1Value := -1000000.0, [0,227].Criteria2Value := -1000000.0, [0,227].ActionValue := -1000000.0, [0,228].Criteria1 := -999, [0,228].Criteria1Operator := -999, [0,228].Boolean := -999, [0,228].Criteria2 := -999, [0,228].Criteria2Operator := -999, [0,228].Action := -999, [0,228].Label := -999, [0,228].Criteria1Value := -1000000.0, [0,228].Criteria2Value := -1000000.0, [0,228].ActionValue := -1000000.0, [0,229].Criteria1 := -999, [0,229].Criteria1Operator := -999, [0,229].Boolean := -999, [0,229].Criteria2 := -999, [0,229].Criteria2Operator := -999, [0,229].Action := -999, [0,229].Label := -999, [0,229].Criteria1Value := -1000000.0, [0,229].Criteria2Value := -1000000.0, [0,229].ActionValue := -1000000.0, [0,230].Criteria1 := -999, [0,230].Criteria1Operator := -999, [0,230].Boolean := -999, [0,230].Criteria2 := -999, [0,230].Criteria2Operator := -999, [0,230].Action := -999, [0,230].Label := -999, [0,230].Criteria1Value := -1000000.0, [0,230].Criteria2Value := -1000000.0, [0,230].ActionValue := -1000000.0, [0,231].Criteria1 := -999, [0,231].Criteria1Operator := -999, [0,231].Boolean := -999, [0,231].Criteria2 := -999, [0,231].Criteria2Operator := -999, [0,231].Action := -999, [0,231].Label := -999, [0,231].Criteria1Value := -1000000.0,
        [0,231].Criteria2Value := -1000000.0, [0,231].ActionValue := -1000000.0, [0,232].Criteria1 := -999, [0,232].Criteria1Operator := -999, [0,232].Boolean := -999, [0,232].Criteria2 := -999, [0,232].Criteria2Operator := -999, [0,232].Action := -999, [0,232].Label := -999, [0,232].Criteria1Value := -1000000.0, [0,232].Criteria2Value := -1000000.0, [0,232].ActionValue := -1000000.0, [0,233].Criteria1 := -999, [0,233].Criteria1Operator := -999, [0,233].Boolean := -999, [0,233].Criteria2 := -999, [0,233].Criteria2Operator := -999, [0,233].Action := -999, [0,233].Label := -999, [0,233].Criteria1Value := -1000000.0, [0,233].Criteria2Value := -1000000.0, [0,233].ActionValue := -1000000.0, [0,234].Criteria1 := -999, [0,234].Criteria1Operator := -999, [0,234].Boolean := -999, [0,234].Criteria2 := -999, [0,234].Criteria2Operator := -999, [0,234].Action := -999, [0,234].Label := -999, [0,234].Criteria1Value := -1000000.0, [0,234].Criteria2Value := -1000000.0, [0,234].ActionValue := -1000000.0, [0,235].Criteria1 := -999, [0,235].Criteria1Operator := -999, [0,235].Boolean := -999, [0,235].Criteria2 := -999, [0,235].Criteria2Operator := -999, [0,235].Action := -999, [0,235].Label := -999, [0,235].Criteria1Value := -1000000.0, [0,235].Criteria2Value := -1000000.0, [0,235].ActionValue := -1000000.0, [0,236].Criteria1 := -999, [0,236].Criteria1Operator := -999, [0,236].Boolean := -999, [0,236].Criteria2 := -999, [0,236].Criteria2Operator := -999, [0,236].Action := -999, [0,236].Label := -999, [0,236].Criteria1Value := -1000000.0, [0,236].Criteria2Value := -1000000.0, [0,236].ActionValue := -1000000.0, [0,237].Criteria1 := -999, [0,237].Criteria1Operator := -999, [0,237].Boolean := -999, [0,237].Criteria2 := -999, [0,237].Criteria2Operator := -999, [0,237].Action := -999, [0,237].Label := -999, [0,237].Criteria1Value := -1000000.0,
        [0,237].Criteria2Value := -1000000.0, [0,237].ActionValue := -1000000.0, [0,238].Criteria1 := -999, [0,238].Criteria1Operator := -999, [0,238].Boolean := -999, [0,238].Criteria2 := -999, [0,238].Criteria2Operator := -999, [0,238].Action := -999, [0,238].Label := -999, [0,238].Criteria1Value := -1000000.0, [0,238].Criteria2Value := -1000000.0, [0,238].ActionValue := -1000000.0, [0,239].Criteria1 := -999, [0,239].Criteria1Operator := -999, [0,239].Boolean := -999, [0,239].Criteria2 := -999, [0,239].Criteria2Operator := -999, [0,239].Action := -999, [0,239].Label := -999, [0,239].Criteria1Value := -1000000.0, [0,239].Criteria2Value := -1000000.0, [0,239].ActionValue := -1000000.0, [0,240].Criteria1 := -999, [0,240].Criteria1Operator := -999, [0,240].Boolean := -999, [0,240].Criteria2 := -999, [0,240].Criteria2Operator := -999, [0,240].Action := -999, [0,240].Label := -999, [0,240].Criteria1Value := -1000000.0, [0,240].Criteria2Value := -1000000.0, [0,240].ActionValue := -1000000.0, [0,241].Criteria1 := -999, [0,241].Criteria1Operator := -999, [0,241].Boolean := -999, [0,241].Criteria2 := -999, [0,241].Criteria2Operator := -999, [0,241].Action := -999, [0,241].Label := -999, [0,241].Criteria1Value := -1000000.0, [0,241].Criteria2Value := -1000000.0, [0,241].ActionValue := -1000000.0, [0,242].Criteria1 := -999, [0,242].Criteria1Operator := -999, [0,242].Boolean := -999, [0,242].Criteria2 := -999, [0,242].Criteria2Operator := -999, [0,242].Action := -999, [0,242].Label := -999, [0,242].Criteria1Value := -1000000.0, [0,242].Criteria2Value := -1000000.0, [0,242].ActionValue := -1000000.0, [0,243].Criteria1 := -999, [0,243].Criteria1Operator := -999, [0,243].Boolean := -999, [0,243].Criteria2 := -999, [0,243].Criteria2Operator := -999, [0,243].Action := -999, [0,243].Label := -999, [0,243].Criteria1Value := -1000000.0,
        [0,243].Criteria2Value := -1000000.0, [0,243].ActionValue := -1000000.0, [0,244].Criteria1 := -999, [0,244].Criteria1Operator := -999, [0,244].Boolean := -999, [0,244].Criteria2 := -999, [0,244].Criteria2Operator := -999, [0,244].Action := -999, [0,244].Label := -999, [0,244].Criteria1Value := -1000000.0, [0,244].Criteria2Value := -1000000.0, [0,244].ActionValue := -1000000.0, [0,245].Criteria1 := -999, [0,245].Criteria1Operator := -999, [0,245].Boolean := -999, [0,245].Criteria2 := -999, [0,245].Criteria2Operator := -999, [0,245].Action := -999, [0,245].Label := -999, [0,245].Criteria1Value := -1000000.0, [0,245].Criteria2Value := -1000000.0, [0,245].ActionValue := -1000000.0, [0,246].Criteria1 := -999, [0,246].Criteria1Operator := -999, [0,246].Boolean := -999, [0,246].Criteria2 := -999, [0,246].Criteria2Operator := -999, [0,246].Action := -999, [0,246].Label := -999, [0,246].Criteria1Value := -1000000.0, [0,246].Criteria2Value := -1000000.0, [0,246].ActionValue := -1000000.0, [0,247].Criteria1 := -999, [0,247].Criteria1Operator := -999, [0,247].Boolean := -999, [0,247].Criteria2 := -999, [0,247].Criteria2Operator := -999, [0,247].Action := -999, [0,247].Label := -999, [0,247].Criteria1Value := -1000000.0, [0,247].Criteria2Value := -1000000.0, [0,247].ActionValue := -1000000.0, [0,248].Criteria1 := -999, [0,248].Criteria1Operator := -999, [0,248].Boolean := -999, [0,248].Criteria2 := -999, [0,248].Criteria2Operator := -999, [0,248].Action := -999, [0,248].Label := -999, [0,248].Criteria1Value := -1000000.0, [0,248].Criteria2Value := -1000000.0, [0,248].ActionValue := -1000000.0, [0,249].Criteria1 := -999, [0,249].Criteria1Operator := -999, [0,249].Boolean := -999, [0,249].Criteria2 := -999, [0,249].Criteria2Operator := -999, [0,249].Action := -999, [0,249].Label := -999, [0,249].Criteria1Value := -1000000.0,
        [0,249].Criteria2Value := -1000000.0, [0,249].ActionValue := -1000000.0, [0,250].Criteria1 := -999, [0,250].Criteria1Operator := -999, [0,250].Boolean := -999, [0,250].Criteria2 := -999, [0,250].Criteria2Operator := -999, [0,250].Action := -999, [0,250].Label := -999, [0,250].Criteria1Value := -1000000.0, [0,250].Criteria2Value := -1000000.0, [0,250].ActionValue := -1000000.0, [1,0].Action := 300701, [1,1].Step := 1, [1,2].Step := 2, [1,2].Action := 700104, [1,2].ActionValue := 1.0, [1,3].Step := 3, [1,3].Action := 800101, [1,3].ActionValue := 1.0, [1,4].Step := 4, [1,4].Criteria1 := 800103, [1,4].Criteria1Operator := 1, [1,4].Boolean := 2, [1,4].Criteria2 := 1100602, [1,4].Criteria2Operator := 1, [1,4].Action := 700104, [1,4].Criteria1Value := 1.0, [1,4].Criteria2Value := 2.0, [1,4].ActionValue := 1.0, [1,5].Step := 5, [1,5].Action := 800101, [1,5].ActionValue := 1.0, [1,6].Step := 6, [1,6].Criteria1 := 800103, [1,6].Criteria1Operator := 1, [1,6].Boolean := 2, [1,6].Criteria2 := 1100602, [1,6].Criteria2Operator := 1, [1,6].Action := 700104, [1,6].Criteria1Value := 1.0, [1,6].Criteria2Value := 2.0, [1,6].ActionValue := 1.0, [1,7].Step := 7, [1,7].Action := 800101, [1,7].ActionValue := 1.0, [1,8].Step := 8, [1,8].Criteria1 := 800103, [1,8].Criteria1Operator := 1, [1,8].Boolean := 2, [1,8].Criteria2 := 1100602, [1,8].Criteria2Operator := 1, [1,8].Action := 700104, [1,8].Criteria1Value := 1.0, [1,8].Criteria2Value := 2.0, [1,8].ActionValue := 1.0, [1,9].Step := 9, [1,9].Action := 1800001, [1,9].ActionValue := 1.0, [1,10].Step := 10,
        [1,10].Action := 1700011, [1,10].ActionValue := 1.0, [1,11].Criteria1 := -999, [1,11].Criteria1Operator := -999, [1,11].Boolean := -999, [1,11].Criteria2 := -999, [1,11].Criteria2Operator := -999, [1,11].Action := -999, [1,11].Label := -999, [1,11].Criteria1Value := -1000000.0, [1,11].Criteria2Value := -1000000.0, [1,11].ActionValue := -1000000.0, [1,12].Criteria1 := -999, [1,12].Criteria1Operator := -999, [1,12].Boolean := -999, [1,12].Criteria2 := -999, [1,12].Criteria2Operator := -999, [1,12].Action := -999, [1,12].Label := -999, [1,12].Criteria1Value := -1000000.0, [1,12].Criteria2Value := -1000000.0, [1,12].ActionValue := -1000000.0, [1,13].Criteria1 := -999, [1,13].Criteria1Operator := -999, [1,13].Boolean := -999, [1,13].Criteria2 := -999, [1,13].Criteria2Operator := -999, [1,13].Action := -999, [1,13].Label := -999, [1,13].Criteria1Value := -1000000.0, [1,13].Criteria2Value := -1000000.0, [1,13].ActionValue := -1000000.0, [1,14].Criteria1 := -999, [1,14].Criteria1Operator := -999, [1,14].Boolean := -999, [1,14].Criteria2 := -999, [1,14].Criteria2Operator := -999, [1,14].Action := -999, [1,14].Label := -999, [1,14].Criteria1Value := -1000000.0, [1,14].Criteria2Value := -1000000.0, [1,14].ActionValue := -1000000.0, [1,15].Criteria1 := -999, [1,15].Criteria1Operator := -999, [1,15].Boolean := -999, [1,15].Criteria2 := -999, [1,15].Criteria2Operator := -999, [1,15].Action := -999, [1,15].Label := -999, [1,15].Criteria1Value := -1000000.0, [1,15].Criteria2Value := -1000000.0, [1,15].ActionValue := -1000000.0, [1,16].Criteria1 := -999, [1,16].Criteria1Operator := -999, [1,16].Boolean := -999, [1,16].Criteria2 := -999, [1,16].Criteria2Operator := -999, [1,16].Action := -999, [1,16].Label := -999, [1,16].Criteria1Value := -1000000.0,
